(* IEC 61131-3 sources: station-control-three-platforms/codesys/src, 8 files *)

(* ---- ST_EvalRecipe.st ---- *)
// Evaluation recipe of FB_CurveEval as one structure. Not in the Siemens original: there the bench
// writes the recipe straight into the multi-instance Station.Eval. CODESYS refuses that
// (C0037 "'Eval' is no input of 'FB_HandleStation'"), so the station takes the recipe by reference
// and copies it into its own evaluation instance when it tares, once per part.
TYPE ST_EvalRecipe :
STRUCT
    Mode : INT := 3;
    GateX : REAL := 3.0;   // mm
    Gate2X : REAL := 10.0;   // mm
    PeakXLo : REAL := 13.0;   // mm
    PeakXHi : REAL := 26.0;   // mm
    StepSpan : REAL := 2.0;   // mm
    StopF : REAL := 30.0;   // N
    G1Lo : REAL;
    G1Hi : REAL;
    MeanLo : REAL;
    MeanHi : REAL;
    HystLo : REAL;
    HystHi : REAL;
    RetFMin : REAL;
    G2Lo : REAL;
    G2Hi : REAL;
    PeakFLo : REAL;
    PeakFHi : REAL;
    PeakXMin : REAL;
    PeakXMax : REAL;
    StepLo : REAL;
    StopXLo : REAL;
    StopXHi : REAL;
    EnvX0 : REAL := 1.0;   // mm
    EnvDx : REAL := 0.5;   // mm
    EnvN : INT := 55;
    EnvLo : ARRAY[0..63] OF REAL;   // N
    EnvHi : ARRAY[0..63] OF REAL;   // N
END_STRUCT
END_TYPE

(* ---- GVL_TestData.st ---- *)
// Generated by tools/testdata.py from siemens/scl/test/DB_TestData.scl. Do not edit.
// Recorded force-travel curves, the evaluation recipe and the expected values of the 14 replay cases.
{attribute 'qualified_only'}
VAR_GLOBAL
    NCurves : INT := 10;
    NCases : INT := 14;
    NSamples : INT := 5932;
    Tol : REAL := 0.001;
    GoodCurve : INT := 0;
    BadCurve : INT := 6;
    GateX : REAL := 3.0;
    Gate2X : REAL := 10.0;
    PeakXLo : REAL := 13.0;
    PeakXHi : REAL := 26.0;
    StepSpan : REAL := 2.0;
    StopF : REAL := 30.0;
    EnvX0 : REAL := 1.0;
    EnvDx : REAL := 0.5;
    EnvN : INT := 55;
    CurveStart : ARRAY[0..15] OF INT := [0, 620, 1246, 1746, 2366, 2988, 3606, 4228, 4728, 5310, 0, 0, 0, 0, 0, 0];
    CurveNPull : ARRAY[0..15] OF INT := [310, 313, 250, 310, 311, 309, 311, 250, 291, 311, 0, 0, 0, 0, 0, 0];
    CaseCurve : ARRAY[1..32] OF INT := [0, 1, 2, 3, 4, 5, 6, 7, 8, 9, 9, 8, 0, 3, 0, 0, 0, 0, 0, 0, 0, 0, 0, 0, 0, 0, 0, 0, 0, 0, 0, 0];
    CaseMode : ARRAY[1..32] OF INT := [3, 3, 3, 3, 3, 3, 3, 3, 3, 3, 2, 1, 4, 4, 0, 0, 0, 0, 0, 0, 0, 0, 0, 0, 0, 0, 0, 0, 0, 0, 0, 0];
    ExpOk : ARRAY[1..32] OF BOOL := [TRUE, TRUE, FALSE, FALSE, FALSE, FALSE, FALSE, FALSE, FALSE, FALSE, TRUE, TRUE, TRUE, TRUE, FALSE, FALSE, FALSE, FALSE, FALSE, FALSE, FALSE, FALSE, FALSE, FALSE, FALSE, FALSE, FALSE, FALSE, FALSE, FALSE, FALSE, FALSE];
    ExpNok : ARRAY[1..32] OF INT := [0, 0, 2, 2, 2, 3, 5, 2, 9, 2, 0, 0, 0, 0, 0, 0, 0, 0, 0, 0, 0, 0, 0, 0, 0, 0, 0, 0, 0, 0, 0, 0];
    ExpEnvViol : ARRAY[1..32] OF INT := [0, 0, 43, 0, 17, 41, 41, 43, 1, 0, 0, 1, 0, 0, 0, 0, 0, 0, 0, 0, 0, 0, 0, 0, 0, 0, 0, 0, 0, 0, 0, 0];
    ExpEnvNodes : ARRAY[1..32] OF INT := [55, 55, 46, 55, 55, 55, 55, 46, 55, 55, 55, 55, 55, 55, 0, 0, 0, 0, 0, 0, 0, 0, 0, 0, 0, 0, 0, 0, 0, 0, 0, 0];
    ExpFeat : ARRAY[0..287] OF REAL := [6.9821014, 5.37568, 6.1788907, 1.6064217, 10.845588, 16.818577, 19.848608, 3.9388027, 29.783041, 7.205183, 5.0210447, 6.113114, 2.1841383, 11.2528515, 17.15133, 18.303595, 4.152199, 30.096466, 4.183258, 2.565676, 3.374467, 1.6175817, 6.124597, 40.227142, 23.940363, 0.0, 23.785864, 5.1918726, 3.556863, 4.3743677, 1.6350094, 9.031395, 14.923322, 19.814, 3.9026327, 29.81065, 4.6947575, 3.0623243, 3.8785408, 1.632433, 8.425375, 14.073351, 19.786457, 3.8736982, 29.815647, 10.499536, 1.8700012, 6.184768, 8.629534, 14.390507, 20.330584, 19.78603, 3.8881645, 29.722036, 7.0127378, 5.3387175, 6.175728, 1.67402, 7.371472, 8.326099, 25.861488, 0.032551765, 29.877676, 4.238579, 2.6031868, 3.420883, 1.6353921, 6.187137, 41.858364, 23.904263, 0.0, 23.727392, 7.0128746, 5.3684235, 6.190649, 1.6444514, 10.856109, 16.749855, 19.791138, 3.8845482, 27.874788, 6.2380857, 2.573432, 4.405759, 3.6646535, 10.107543, 15.954138, 19.8363, 3.8773146, 29.792097, 6.2380857, 2.573432, 4.405759, 3.6646535, 10.107543, 15.954138, 19.8363, 3.8773146, 29.792097, 7.0128746, 5.3684235, 6.190649, 1.6444514, 10.856109, 16.749855, 19.791138, 3.8845482, 27.874788, 6.9821014, 5.37568, 6.1788907, 1.6064217, 10.845588, 16.818577, 19.848608, 3.9388027, 29.783041, 5.1918726, 3.556863, 4.3743677, 1.6350094, 9.031395, 14.923322, 19.814, 3.9026327, 29.81065, 0.0, 0.0, 0.0, 0.0, 0.0, 0.0, 0.0, 0.0, 0.0, 0.0, 0.0, 0.0, 0.0, 0.0, 0.0, 0.0, 0.0, 0.0, 0.0, 0.0, 0.0, 0.0, 0.0, 0.0, 0.0, 0.0, 0.0, 0.0, 0.0, 0.0, 0.0, 0.0, 0.0, 0.0, 0.0, 0.0, 0.0, 0.0, 0.0, 0.0, 0.0, 0.0, 0.0, 0.0, 0.0, 0.0, 0.0, 0.0, 0.0, 0.0, 0.0, 0.0, 0.0, 0.0, 0.0, 0.0, 0.0, 0.0, 0.0, 0.0, 0.0, 0.0, 0.0, 0.0, 0.0, 0.0, 0.0, 0.0, 0.0, 0.0, 0.0, 0.0, 0.0, 0.0, 0.0, 0.0, 0.0, 0.0, 0.0, 0.0, 0.0, 0.0, 0.0, 0.0, 0.0, 0.0, 0.0, 0.0, 0.0, 0.0, 0.0, 0.0, 0.0, 0.0, 0.0, 0.0, 0.0, 0.0, 0.0, 0.0, 0.0, 0.0, 0.0, 0.0, 0.0, 0.0, 0.0, 0.0, 0.0, 0.0, 0.0, 0.0, 0.0, 0.0, 0.0, 0.0, 0.0, 0.0, 0.0, 0.0, 0.0, 0.0, 0.0, 0.0, 0.0, 0.0, 0.0, 0.0, 0.0, 0.0, 0.0, 0.0, 0.0, 0.0, 0.0, 0.0, 0.0, 0.0, 0.0, 0.0, 0.0, 0.0, 0.0, 0.0, 0.0, 0.0, 0.0, 0.0, 0.0, 0.0, 0.0, 0.0, 0.0, 0.0, 0.0, 0.0, 0.0, 0.0, 0.0, 0.0, 0.0, 0.0];
    ExpFeatValid : ARRAY[0..287] OF BOOL := [TRUE, TRUE, TRUE, TRUE, TRUE, TRUE, TRUE, TRUE, TRUE, TRUE, TRUE, TRUE, TRUE, TRUE, TRUE, TRUE, TRUE, TRUE, TRUE, TRUE, TRUE, TRUE, TRUE, TRUE, TRUE, TRUE, TRUE, TRUE, TRUE, TRUE, TRUE, TRUE, TRUE, TRUE, TRUE, TRUE, TRUE, TRUE, TRUE, TRUE, TRUE, TRUE, TRUE, TRUE, TRUE, TRUE, TRUE, TRUE, TRUE, TRUE, TRUE, TRUE, TRUE, TRUE, TRUE, TRUE, TRUE, TRUE, TRUE, TRUE, TRUE, TRUE, TRUE, TRUE, TRUE, TRUE, TRUE, TRUE, TRUE, TRUE, TRUE, TRUE, TRUE, TRUE, TRUE, TRUE, TRUE, TRUE, TRUE, TRUE, TRUE, TRUE, TRUE, TRUE, TRUE, TRUE, TRUE, TRUE, TRUE, TRUE, TRUE, TRUE, TRUE, TRUE, TRUE, TRUE, TRUE, TRUE, TRUE, TRUE, TRUE, TRUE, TRUE, TRUE, TRUE, TRUE, TRUE, TRUE, TRUE, TRUE, TRUE, TRUE, TRUE, TRUE, TRUE, TRUE, TRUE, TRUE, TRUE, TRUE, TRUE, TRUE, TRUE, TRUE, TRUE, TRUE, FALSE, FALSE, FALSE, FALSE, FALSE, FALSE, FALSE, FALSE, FALSE, FALSE, FALSE, FALSE, FALSE, FALSE, FALSE, FALSE, FALSE, FALSE, FALSE, FALSE, FALSE, FALSE, FALSE, FALSE, FALSE, FALSE, FALSE, FALSE, FALSE, FALSE, FALSE, FALSE, FALSE, FALSE, FALSE, FALSE, FALSE, FALSE, FALSE, FALSE, FALSE, FALSE, FALSE, FALSE, FALSE, FALSE, FALSE, FALSE, FALSE, FALSE, FALSE, FALSE, FALSE, FALSE, FALSE, FALSE, FALSE, FALSE, FALSE, FALSE, FALSE, FALSE, FALSE, FALSE, FALSE, FALSE, FALSE, FALSE, FALSE, FALSE, FALSE, FALSE, FALSE, FALSE, FALSE, FALSE, FALSE, FALSE, FALSE, FALSE, FALSE, FALSE, FALSE, FALSE, FALSE, FALSE, FALSE, FALSE, FALSE, FALSE, FALSE, FALSE, FALSE, FALSE, FALSE, FALSE, FALSE, FALSE, FALSE, FALSE, FALSE, FALSE, FALSE, FALSE, FALSE, FALSE, FALSE, FALSE, FALSE, FALSE, FALSE, FALSE, FALSE, FALSE, FALSE, FALSE, FALSE, FALSE, FALSE, FALSE, FALSE, FALSE, FALSE, FALSE, FALSE, FALSE, FALSE, FALSE, FALSE, FALSE, FALSE, FALSE, FALSE, FALSE, FALSE, FALSE, FALSE, FALSE, FALSE, FALSE, FALSE, FALSE, FALSE, FALSE, FALSE, FALSE, FALSE, FALSE, FALSE, FALSE, FALSE, FALSE, FALSE, FALSE, FALSE, FALSE, FALSE, FALSE, FALSE, FALSE, FALSE, FALSE];
    Lim : ARRAY[0..63] OF REAL := [0.0, 0.0, 0.0, 0.0, 0.0, 0.0, 0.0, 0.0, 0.0, 15.241609, 18.417305, 0.0, 0.0, 0.0, 0.0, 0.0, 5.896105, 8.38203, 0.0, 0.0, 0.0, 0.0, 0.0, 9.4181, 12.402887, 14.982571, 18.676344, 17.139359, 22.516165, 2.9451215, 28.690018, 30.871372, 0.0, 0.0, 5.186474, 7.2080727, -0.5455249, 3.975223, 1.0, 9.212741, 12.608247, 14.728432, 18.930483, 16.769424, 22.886099, 2.8110514, 28.539938, 31.021452, 0.0, 0.0, 0.0, 0.0, 0.0, 0.0, 0.0, 0.0, 0.0, 0.0, 0.0, 0.0, 0.0, 0.0, 0.0, 0.0];
    EnvLo : ARRAY[0..63] OF REAL := [4.5024867, 4.5624857, 4.530773, 4.5635424, 4.573186, 4.617667, 4.6239376, 4.670679, 4.725596, 4.700003, 4.8820324, 4.926072, 5.163019, 5.6595745, 7.878658, 8.020163, 8.08159, 8.207902, 8.30263, 8.350869, 8.425625, 8.550419, 8.607436, 8.764787, 8.845735, 8.9147835, 8.99205, 9.068602, 9.331687, 9.416069, 9.513143, 9.665618, 10.123489, 10.642103, 11.14989, 11.027167, 10.830289, 10.428676, 10.27112, 10.313659, 10.363278, 10.468162, 10.585302, 10.677869, 10.748317, 10.8695135, 10.998811, 11.099038, 11.214338, 11.278554, 11.41541, 11.506263, 11.623229, 11.713954, 11.844806, 0.0, 0.0, 0.0, 0.0, 0.0, 0.0, 0.0, 0.0, 0.0];
    EnvHi : ARRAY[0..63] OF REAL := [9.917023, 9.98225, 9.992803, 10.004515, 10.029344, 10.026862, 10.070514, 10.102605, 12.041139, 12.557893, 12.779339, 12.91771, 13.360822, 13.471234, 13.533369, 13.642666, 13.729599, 13.860825, 13.911284, 13.990431, 14.0966015, 14.182879, 14.296827, 14.390328, 14.4539795, 14.551714, 14.698472, 15.185006, 15.688478, 16.23098, 16.795422, 17.309069, 17.854668, 18.362646, 18.931261, 18.921373, 19.396362, 19.986576, 19.496552, 19.897247, 19.346785, 18.766773, 16.553541, 16.354622, 16.457827, 16.512941, 16.617954, 16.769545, 16.847044, 16.997396, 17.054838, 17.213253, 17.348417, 17.397055, 17.536877, 0.0, 0.0, 0.0, 0.0, 0.0, 0.0, 0.0, 0.0, 0.0];
    X : ARRAY[0..5931] OF REAL := [0.0, -0.0033742767, 0.10472685, 0.19745024, 0.29981726, 0.39700347, 0.49491304, 0.6008226, 0.6972801, 0.7991843, 0.90281725, 0.99573755, 1.0995567, 1.1978173, 1.2951844, 1.3980939, 1.4998226, 1.5985514, 1.7018226, 1.8003706, 1.8912854, 1.999562, 2.0993705, 2.1909237, 2.2984662, 2.3891046, 2.4932854, 2.601009, 2.6959238, 2.796014, 2.894743, 2.9955568, 3.092743, 3.1978333, 3.292743, 3.3987377, 3.4987428, 3.59511, 3.6955674, 3.7989292, 3.8956633, 3.9927535, 4.0977483, 4.197296, 4.292573, 4.399477, 4.4931207, 4.593658, 4.6908493, 4.7944875, 4.8961205, 4.9969397, 5.094764, 5.18994, 5.2910357, 5.394844, 5.489573, 5.5893974, 5.6894984, 5.7891207, 5.893126, 5.989312, 6.076935, 6.1627493, 6.2443776, 6.328378, 6.4094586, 6.5168147, 6.6171765, 6.718815, 6.8094583, 6.9220915, 7.0171022, 7.1126394, 7.213565, 7.3112035, 7.4117403, 7.511751, 7.606661, 7.708384, 7.81248, 7.9090276, 8.005486, 8.110033, 8.2134, 8.307496, 8.410586, 8.505591, 8.600773, 8.702959, 8.809416, 8.908698, 8.999699, 9.103602, 9.201704, 9.301433, 9.39789, 9.503613, 9.601155, 9.699528, 9.802805, 9.89989, 10.003895, 10.098449, 10.201262, 10.298172, 10.399454, 10.497454, 10.592826, 10.699917, 10.798554, 10.89847, 10.996193, 11.098837, 11.192114, 11.287757, 11.391119, 11.496119, 11.592933, 11.693028, 11.786496, 11.891943, 11.991592, 12.0868635, 12.186582, 12.291321, 12.380411, 12.48514, 12.584327, 12.683965, 12.787603, 12.888337, 12.989885, 13.08306, 13.187704, 13.284523, 13.3848, 13.487896, 13.587353, 13.678811, 13.784454, 13.882715, 13.981008, 14.078545, 14.183087, 14.28164, 14.38038, 14.475013, 14.574927, 14.682922, 14.780104, 14.878199, 14.975023, 15.076039, 15.17287, 15.271434, 15.363907, 15.460098, 15.557104, 15.660487, 15.751045, 15.851062, 15.951705, 16.053541, 16.149647, 16.244019, 16.34385, 16.440685, 16.537062, 16.62862, 16.734083, 16.83637, 16.92229, 17.019585, 17.119505, 17.217972, 17.316803, 17.418, 17.508282, 17.611292, 17.70858, 17.800692, 17.902872, 17.99408, 18.09909, 18.191565, 18.287483, 18.387772, 18.49033, 18.585798, 18.676447, 18.777182, 18.874111, 18.979118, 19.070032, 19.165964, 19.270985, 19.360996, 19.462011, 19.55457, 19.65848, 19.755777, 19.848608, 19.970793, 20.087416, 20.211292, 20.32783, 20.445093, 20.557806, 20.648077, 20.741636, 20.84809, 20.953089, 21.043913, 21.147093, 21.24119, 21.348913, 21.449648, 21.545195, 21.634748, 21.745749, 21.841301, 21.946121, 22.040205, 22.143402, 22.240217, 22.341042, 22.44068, 22.53859, 22.634499, 22.738136, 22.838509, 22.941322, 23.042967, 23.129976, 23.239418, 23.335434, 23.430067, 23.531801, 23.641802, 23.734535, 23.835356, 23.933903, 24.02927, 24.133179, 24.232546, 24.332918, 24.43128, 24.52801, 24.624918, 24.728653, 24.823557, 24.925116, 25.026297, 25.123116, 25.230398, 25.325674, 25.426765, 25.523584, 25.621408, 25.71895, 25.820227, 25.919882, 26.019594, 26.116701, 26.216702, 26.315063, 26.42161, 26.524881, 26.622345, 26.714718, 26.815802, 26.917803, 27.014627, 27.115812, 27.214813, 27.312366, 27.413908, 27.51119, 27.612286, 27.709558, 27.811739, 27.911112, 28.007027, 28.111387, 28.199669, 28.301207, 28.40676, 28.508398, 28.60403, 28.701595, 28.8095, 28.900776, 29.00051, 29.101877, 29.200064, 29.301426, 29.398798, 29.500973, 29.572319, 29.6092, 29.646812, 29.686869, 29.716297, 29.758177, 29.799242, 29.837845, 29.867996, 29.91243, 29.94758, 29.943314, 29.928886, 29.886644, 29.850302, 29.813248, 29.77291, 29.739481, 29.693878, 29.666807, 29.625662, 29.588596, 29.545658, 29.446291, 29.346828, 29.248291, 29.144827, 29.049004, 28.937727, 28.847637, 28.75453, 28.642721, 28.549807, 28.448168, 28.348167, 28.251705, 28.151072, 28.05543, 27.9487, 27.857418, 27.751062, 27.654417, 27.556412, 27.45969, 27.360954, 27.257498, 27.15513, 27.059216, 26.958311, 26.85785, 26.761482, 26.654758, 26.5573, 26.460743, 26.360561, 26.257103, 26.160013, 26.06664, 25.96328, 25.863731, 25.76454, 25.668083, 25.56563, 25.464897, 25.367987, 25.26344, 25.167982, 25.070257, 24.966524, 24.871796, 24.767876, 24.67279, 24.576056, 24.471146, 24.368502, 24.26669, 24.170046, 24.073677, 23.97786, 23.87113, 23.777668, 23.676853, 23.576395, 23.480204, 23.375023, 23.272934, 23.17702, 23.081102, 22.978556, 22.88028, 22.779646, 22.677635, 22.582449, 22.482183, 22.376087, 22.28681, 22.185173, 22.084444, 21.981167, 21.891161, 21.780619, 21.684343, 21.589523, 21.48388, 21.391508, 21.285975, 21.187326, 21.08787, 20.986044, 20.88931, 20.790411, 20.692492, 20.591034, 20.4904, 20.394842, 20.293018, 20.197294, 20.102022, 19.994108, 19.893831, 19.797018, 19.694916, 19.590475, 19.501102, 19.397188, 19.298725, 19.19691, 19.100178, 18.99881, 18.902714, 18.797997, 18.700708, 18.604261, 18.502884, 18.39889, 18.303162, 18.206156, 18.103241, 17.99897, 17.907688, 17.802235, 17.704773, 17.608416, 17.508411, 17.407219, 17.30849, 17.209394, 17.109943, 17.011847, 16.906948, 16.809395, 16.708118, 16.613565, 16.507107, 16.412107, 16.31701, 16.208832, 16.112278, 16.011374, 15.918001, 15.814639, 15.7179, 15.617182, 15.515448, 15.413996, 15.3189, 15.21989, 15.117075, 15.018708, 14.91516, 14.81798, 14.721788, 14.619889, 14.519878, 14.4160595, 14.324873, 14.220602, 14.128693, 14.019857, 13.914687, 13.827314, 13.7215, 13.626677, 13.521501, 13.424581, 13.327847, 13.228756, 13.133394, 13.029112, 12.930293, 12.828841, 12.727287, 12.62883, 12.531464, 12.429921, 12.327181, 12.229639, 12.131453, 12.032723, 11.925458, 11.833815, 11.732442, 11.633894, 11.536803, 11.433075, 11.328346, 11.23716, 11.135245, 11.032245, 10.939425, 10.837878, 10.737963, 10.632873, 10.537234, 10.437139, 10.339868, 10.24041, 10.143681, 10.045037, 9.939037, 9.833128, 9.744676, 9.642303, 9.540303, 9.441941, 9.343032, 9.2415695, 9.141931, 9.047192, 8.943649, 8.843558, 8.747462, 8.645282, 8.554914, 8.446638, 8.344186, 8.247452, 8.145633, 8.051356, 7.9505424, 7.854803, 7.749255, 7.6534357, 7.5542603, 7.453893, 7.3493347, 7.2504253, 7.1519732, 7.054606, 6.9581485, 6.8538775, 6.7531433, 6.657409, 6.5563293, 6.4607816, 6.3632812, 6.274286, 6.1935673, 6.108753, 6.03021, 5.9339066, 5.8310876, 5.731545, 5.6369066, 5.531364, 5.437353, 5.337811, 5.2275395, 5.126901, 5.03872, 4.9384384, 4.8375287, 4.739082, 4.634901, 4.5331616, 4.4404383, 4.329167, 4.233348, 4.1344438, 4.0365286, 3.9392576, 3.834167, 3.7369862, 3.633433, 3.5345287, 3.4394383, 3.3372576, 3.2332575, 3.140433, 3.043066, 2.9320712, 2.8413372, 2.7396085, 2.6366086, 2.5347893, 2.441518, 2.342518, 2.2378001, 2.1382415, 2.034066, 1.9376031, 1.8358798, 1.7395127, 1.6385127, 1.540151, 1.4401511, 1.3368851, 1.2400553, 1.133151, 1.0449648, 0.939784, 0.8416882, 0.7337893, 0.6410499, 0.5402415, 0.43896484, 0.34032118, 0.23696484, 0.14223076, 0.03723076, 0.07943374, 0.0, 0.058969617, 0.1601451, 0.25842172, 0.36087385, 0.45877805, 0.5548792, 0.6574271, 0.75815046, 0.85487384, 0.9517888, 1.053975, 1.1582409, 1.2541559, 1.3572463, 1.4556025, 1.5523367, 1.6556187, 1.7556983, 1.8526186, 1.9547037, 2.0571558, 2.1517036, 2.2567995, 2.3577092, 2.4552517, 2.5556185, 2.6554377, 2.7547994, 2.850161, 2.9497144, 3.0517995, 3.1496186, 3.257076, 3.3558953, 3.4521666, 3.5518048, 3.653624, 3.7534378, 3.852991, 3.9552622, 4.04972, 4.1526294, 4.255996, 4.3528047, 4.4510016, 4.5480866, 4.6492677, 4.7482677, 4.853805, 4.9477253, 5.051906, 5.151358, 5.2348957, 5.3198113, 5.4007053, 5.4895253, 5.573419, 5.673228, 5.771866, 5.871143, 5.969329, 6.072978, 6.165616, 6.2763395, 6.37834, 6.4693394, 6.5714407, 6.6652493, 6.770627, 6.8630843, 6.9633555, 7.0697227, 7.168909, 7.2685523, 7.3637385, 7.4669037, 7.563648, 7.6645527, 7.7610154, 7.8674674, 7.9631057, 8.063478, 8.159749, 8.254574, 8.355664, 8.462856, 8.553574, 8.662393, 8.762766, 8.8588505, 8.952951, 9.056047, 9.15259, 9.251148, 9.357691, 9.453968, 9.555329, 9.654702, 9.75134, 9.855978, 9.954888, 10.04817, 10.15099, 10.252255, 10.3547125, 10.451904, 10.551271, 10.646809, 10.748909, 10.853186, 10.952457, 11.050553, 11.14801, 11.246378, 11.350468, 11.444835, 11.546383, 11.644745, 11.748659, 11.844665, 11.942393, 12.038213, 12.13958, 12.245122, 12.339048, 12.439409, 12.540957, 12.639862, 12.740053, 12.837516, 12.932607, 13.040059, 13.139059, 13.238154, 13.338431, 13.4359, 13.5304575, 13.635559, 13.72675, 13.818857, 13.918681, 14.016246, 14.117352, 14.217459, 14.311023, 14.407762, 14.50431, 14.610332, 14.701975, 14.796544, 14.899007, 14.994475, 15.085858, 15.194316, 15.28988, 15.3827095, 15.478273, 15.579289, 15.676763, 15.776773, 15.875156, 15.973704, 16.068811, 16.163736, 16.2553, 16.359764, 16.457323, 16.552242, 16.653168, 16.743004, 16.841015, 16.939758, 17.037136, 17.140327, 17.235802, 17.331541, 17.428104, 17.52593, 17.631126, 17.718876, 17.81943, 17.915802, 18.00819, 18.111834, 18.202488, 18.303595, 18.407286, 18.52944, 18.65905, 18.7763, 18.901001, 19.0094, 19.106045, 19.20614, 19.303415, 19.40779, 19.507235, 19.609697, 19.70224, 19.802341, 19.900156, 20.002895, 20.102533, 20.202618, 20.304895, 20.402363, 20.497267, 20.599997, 20.69355, 20.796188, 20.893097, 20.992193, 21.097012, 21.191204, 21.29547, 21.400927, 21.492119, 21.598661, 21.689854, 21.794113, 21.885592, 21.988316, 22.08878, 22.190773, 22.293049, 22.38805, 22.484604, 22.585506, 22.687784, 22.784433, 22.885614, 22.98833, 23.082354, 23.185162, 23.283348, 23.381716, 23.482725, 23.583992, 23.68372, 23.78337, 23.879997, 23.972647, 24.07764, 24.179012, 24.279741, 24.376842, 24.48021, 24.577572, 24.6793, 24.773943, 24.874945, 24.974407, 25.07404, 25.175955, 25.274588, 25.366964, 25.468056, 25.566055, 25.66897, 25.770609, 25.869247, 25.965885, 26.0708, 26.170258, 26.2708, 26.36344, 26.460264, 26.56645, 26.666822, 26.763725, 26.867178, 26.958647, 27.05411, 27.163929, 27.263475, 27.364023, 27.460024, 27.559578, 27.659397, 27.761215, 27.85913, 27.956684, 28.054413, 28.157417, 28.249779, 28.357328, 28.453423, 28.551237, 28.653881, 28.746983, 28.850885, 28.955158, 29.047626, 29.149813, 29.249632, 29.350636, 29.44836, 29.546822, 29.64455, 29.74519, 29.845291, 29.898531, 29.932146, 29.975742, 30.014538, 30.052784, 30.09384, 30.124363, 30.161966, 30.199852, 30.23428, 30.276073, 30.279707, 30.259258, 30.220552, 30.182497, 30.147161, 30.109282, 30.07712, 30.027245, 29.995913, 29.958479, 29.921057, 29.88163, 29.803432, 29.702337, 29.604788, 29.508512, 29.404512, 29.309692, 29.208055, 29.105412, 29.010315, 28.907495, 28.810219, 28.708496, 28.606033, 28.511213, 28.409018, 28.308836, 28.206108, 28.11083, 28.009554, 27.920464, 27.817097, 27.714096, 27.614098, 27.519081, 27.421623, 27.311539, 27.215809, 27.113165, 27.011442, 26.923613, 26.819523, 26.72316, 26.624512, 26.518154, 26.424501, 26.324501, 26.223682, 26.12832, 26.023682, 25.925581, 25.826756, 25.725304, 25.633213, 25.526209, 25.431484, 25.327932, 25.231379, 25.124107, 25.027378, 24.92774, 24.827005, 24.72682, 24.634266, 24.533634, 24.435629, 24.333357, 24.235714, 24.134075, 24.037159, 23.934883, 23.83689, 23.733522, 23.644058, 23.538336, 23.439335, 23.337143, 23.241873, 23.141325, 23.039495, 22.943308, 22.836676, 22.740585, 22.643122, 22.548845, 22.443756, 22.34893, 22.245022, 22.14148, 22.045925, 21.948095, 21.845825, 21.747463, 21.648638, 21.544724, 21.452633, 21.34591, 21.252352, 21.149809, 21.053707, 20.957075, 20.850708, 20.75434, 20.64933, 20.556244, 20.450605, 20.35551, 20.255686, 20.158957, 20.061596, 19.960772, 19.857952, 19.762127, 19.659489, 19.561398, 19.463669, 19.359297, 19.259573, 19.161749, 19.060844, 18.962467, 18.862371, 18.765282, 18.660913, 18.566366, 18.460653, 18.360914, 18.270807, 18.172451, 18.065079, 17.969627, 17.871622, 17.768164, 17.67243, 17.567436, 17.47643, 17.368792, 17.271786, 17.17751, 17.071148, 16.969872, 16.872866, 16.770239, 16.681765, 16.574047, 16.477217, 16.370668, 16.275764, 16.177212, 16.073658, 15.979759, 15.87902, 15.777563, 15.671382, 15.586376, 15.481924, 15.379919, 15.276377, 15.181281, 15.08636, 14.982185, 14.887541, 14.778909, 14.685083, 14.590627, 14.482345, 14.385892, 14.288073, 14.186977, 14.087796, 13.983977, 13.882429, 13.788419, 13.691237, 13.585786, 13.489599, 13.390775, 13.289956, 13.196493, 13.09286, 12.993312, 12.887945, 12.791126, 12.695663, 12.598573, 12.4952965, 12.398929, 12.295924, 12.19511, 12.095748, 11.997562, 11.899285, 11.795099, 11.700924, 11.59928, 11.501275, 11.400998, 11.296269, 11.20136, 11.098631, 10.997439, 10.901258, 10.802343, 10.704705, 10.604073, 10.503344, 10.405062, 10.304508, 10.20687, 10.110237, 10.015503, 9.908232, 9.80387, 9.70986, 9.613317, 9.510488, 9.412759, 9.315125, 9.2118435, 9.115025, 9.007386, 8.917743, 8.812657, 8.711567, 8.614014, 8.5132, 8.413094, 8.316461, 8.2181835, 8.115466, 8.0167265, 7.91754, 7.821811, 7.720806, 7.614529, 7.5185294, 7.415439, 7.320343, 7.2262526, 7.1214337, 7.015976, 6.92479, 6.824875, 6.7247844, 6.624508, 6.5194283, 6.4205985, 6.325327, 6.2258644, 6.1244917, 6.02304, 5.9274974, 5.825758, 5.7219496, 5.6314015, 5.536194, 5.44547, 5.3669214, 5.285751, 5.202383, 5.105436, 5.006702, 4.9036064, 4.806521, 4.706877, 4.6049786, 4.5074253, 4.4004254, 4.30834, 4.207973, 4.1086006, 4.004883, 3.9012392, 3.8079624, 3.7125103, 3.6096008, 3.5041487, 3.413053, 3.30342, 3.21142, 3.1053243, 3.0126913, 2.9129572, 2.8093243, 2.699053, 2.6135051, 2.506138, 2.4069571, 2.3082337, 2.2100475, 2.1109626, 2.00642, 1.910505, 1.8110476, 1.7060529, 1.6115955, 1.5136752, 1.4113135, 1.3050423, 1.2158561, 1.1087602, 1.0117602, 0.9073135, 0.8141273, 0.7076752, 0.6063986, 0.50649434, 0.40968055, 0.31476563, 0.20966984, 0.11121774, 0.008217737, 0.0, 0.08626114, 0.16408622, 0.25262398, 0.34693274, 0.44683695, 0.5450178, 0.64548063, 0.7489327, 0.841486, 0.944571, 1.047401, 1.1493956, 1.2461296, 1.3409435, 1.4471296, 1.5429435, 1.6451297, 1.7413158, 1.8395978, 1.9470446, 2.046316, 2.141688, 2.2395074, 2.3439596, 2.440784, 2.540598, 2.6418743, 2.7417786, 2.8391511, 2.9425128, 3.0404222, 3.1325235, 3.2412467, 3.3387947, 3.4342575, 3.5342574, 3.6396246, 3.7380767, 3.8398108, 3.9381723, 4.034534, 4.13063, 4.2379065, 4.332268, 4.4399066, 4.5368214, 4.628816, 4.735364, 4.836087, 4.928742, 5.0387416, 5.130109, 5.239098, 5.3370132, 5.43438, 5.5339227, 5.6311035, 5.731024, 5.8305664, 5.924747, 6.027933, 6.1294813, 6.2354865, 6.3234863, 6.43004, 6.530306, 6.6274014, 6.7249546, 6.8309493, 6.9234123, 7.0274973, 7.1264067, 7.2263165, 7.329322, 7.422141, 7.5283217, 7.6280613, 7.7241464, 7.820609, 7.923875, 8.022885, 8.123976, 8.231061, 8.323157, 8.426066, 8.522167, 8.62453, 8.719806, 8.822077, 8.918812, 9.018099, 9.116663, 9.21195, 9.308865, 9.403785, 9.504344, 9.603817, 9.694104, 9.796387, 9.90503, 9.994046, 10.088147, 10.185254, 10.283903, 10.380095, 10.480473, 10.572754, 10.679222, 10.772696, 10.870611, 10.970898, 11.067276, 11.16219, 11.261116, 11.365132, 11.458878, 11.550426, 11.658532, 11.751276, 11.844559, 11.944931, 12.048128, 12.144404, 12.240521, 12.341804, 12.436001, 12.537735, 12.632028, 12.722315, 12.822873, 12.918155, 13.020804, 13.11182, 13.215831, 13.312203, 13.411315, 13.506406, 13.602703, 13.704895, 13.813751, 13.936825, 14.052898, 14.177792, 14.293041, 14.399817, 14.500093, 14.601089, 14.699647, 14.798828, 14.900009, 14.99928, 15.095919, 15.194653, 15.2962055, 15.402014, 15.493297, 15.597206, 15.696291, 15.793211, 15.894573, 15.994216, 16.094482, 16.197584, 16.296854, 16.395493, 16.494854, 16.593866, 16.69186, 16.793776, 16.89269, 16.994047, 17.094774, 17.193243, 17.292328, 17.389967, 17.489605, 17.591696, 17.690153, 17.79379, 17.88644, 17.984615, 18.091429, 18.188078, 18.289797, 18.389711, 18.487074, 18.585089, 18.683716, 18.787716, 18.88736, 18.982813, 19.084908, 19.180637, 19.287733, 19.378914, 19.481653, 19.58519, 19.688015, 19.784105, 19.885105, 19.981941, 20.080477, 20.177025, 20.277748, 20.381495, 20.474669, 20.585121, 20.684946, 20.782211, 20.869228, 20.983856, 21.075409, 21.175041, 21.27759, 21.37559, 21.48168, 21.57587, 21.669786, 21.769611, 21.87778, 21.970972, 22.07425, 22.1737, 22.27034, 22.372978, 22.464525, 22.568436, 22.673801, 22.76935, 22.873451, 22.968447, 23.068174, 23.167181, 23.262638, 23.363457, 23.448547, 23.490519, 23.525759, 23.558645, 23.595072, 23.638952, 23.6792, 23.715626, 23.748682, 23.789104, 23.828627, 23.864237, 23.902477, 23.940363, 23.9459, 23.91903, 23.88006, 23.848814, 23.799929, 23.76615, 23.732264, 23.693836, 23.654856, 23.61289, 23.575373, 23.54095, 23.499975, 23.465818, 23.40177, 23.306679, 23.211945, 23.113216, 23.009312, 22.915482, 22.810843, 22.714844, 22.607939, 22.5082, 22.41111, 22.315023, 22.216562, 22.114561, 22.017641, 21.91356, 21.818556, 21.71846, 21.61546, 21.519827, 21.423178, 21.322727, 21.2219, 21.118635, 21.017353, 20.921162, 20.821173, 20.717806, 20.617353, 20.519167, 20.423529, 20.323885, 20.222248, 20.122982, 20.017609, 19.922152, 19.82279, 19.728874, 19.628683, 19.527231, 19.420507, 19.328598, 19.226055, 19.12614, 19.027859, 18.92413, 18.830034, 18.725492, 18.621853, 18.528305, 18.429848, 18.329391, 18.231758, 18.133385, 18.02812, 17.93539, 17.828562, 17.731556, 17.632019, 17.53247, 17.435652, 17.331741, 17.23164, 17.13119, 17.039188, 16.934822, 16.834013, 16.72946, 16.632635, 16.541449, 16.433624, 16.337263, 16.238619, 16.140078, 16.041264, 15.936167, 15.837439, 15.731354, 15.643433, 15.542253, 15.437524, 15.340157, 15.234438, 15.1426935, 15.038332, 14.945151, 14.839055, 14.736237, 14.64305, 14.54605, 14.445321, 14.343502, 14.241587, 14.14296, 14.043225, 13.940954, 13.848028, 13.748943, 13.649853, 13.5404005, 13.445395, 13.346565, 13.251119, 13.149114, 13.047938, 12.949023, 12.845475, 12.744108, 12.648922, 12.546831, 12.443922, 12.351374, 12.2532835, 12.144917, 12.04564, 11.948273, 11.850539, 11.755182, 11.652087, 11.552539, 11.4536295, 11.353901, 11.25381, 11.150906, 11.051443, 10.959076, 10.856342, 10.759076, 10.655523, 10.555251, 10.460879, 10.356331, 10.25497, 10.159789, 10.060602, 9.955512, 9.858231, 9.758411, 9.658512, 9.55823, 9.461773, 9.35714, 9.258135, 9.159677, 9.060767, 8.962858, 8.86222, 8.762124, 8.663587, 8.565485, 8.465938, 8.362666, 8.270204, 8.161209, 8.063927, 7.969384, 7.865379, 7.757927, 7.661746, 7.571554, 7.4681025, 7.373012, 7.262645, 7.166826, 7.067826, 6.965905, 6.872453, 6.765549, 6.6689053, 6.567815, 6.467815, 6.374448, 6.27481, 6.170256, 6.0742564, 5.970443, 5.867533, 5.775799, 5.669251, 5.576607, 5.4744263, 5.37507, 5.274251, 5.173602, 5.0736976, 4.973969, 4.87824, 4.7821445, 4.680597, 4.5706925, 4.4696817, 4.3800435, 4.268049, 4.172134, 4.080586, 3.9725008, 3.8796763, 3.7860382, 3.6812189, 3.5841231, 3.479304, 3.376038, 3.285123, 3.1766655, 3.0816603, 2.9889317, 2.8742027, 2.7805698, 2.6814742, 2.58474, 2.4808357, 2.3843784, 2.2894688, 2.1821017, 2.0858252, 1.9848198, 1.8824581, 1.7823783, 1.689091, 1.5809155, 1.4890857, 1.3824581, 1.2849952, 1.1856335, 1.0859048, 0.9898941, 0.8930803, 0.7830696, 0.6876282, 0.5891654, 0.48952705, 0.39324507, 0.29234084, 0.20517014, 0.11862703, 0.044536024, 0.0, 0.059942853, 0.15758651, 0.25440568, 0.3589482, 0.46004933, 0.5611344, 0.6548631, 0.75676733, 0.86150146, 0.95358115, 1.0613099, 1.1569589, 1.2548631, 1.3582249, 1.4564961, 1.5571398, 1.6575068, 1.7561344, 1.8561398, 1.9555973, 2.055959, 2.15731, 2.2549536, 2.355693, 2.4565973, 2.5547833, 2.653778, 2.7529643, 2.8573205, 2.9499643, 3.0485973, 3.154326, 3.258145, 3.3519697, 3.4530602, 3.5616877, 3.6537888, 3.7530653, 3.8539696, 3.9496984, 4.048975, 4.15506, 4.2600656, 4.3559694, 4.450241, 4.553613, 4.6583314, 4.7553368, 4.8541613, 4.952624, 5.0506186, 5.1556134, 5.2568846, 5.3572516, 5.4571557, 5.5487146, 5.6542516, 5.7500815, 5.848257, 5.946342, 6.0442944, 6.131662, 6.2118382, 6.2960143, 6.375015, 6.475398, 6.5699406, 6.673946, 6.7746744, 6.876488, 6.9773183, 7.0665946, 7.1729617, 7.27168, 7.3722386, 7.4740577, 7.5736055, 7.6791425, 7.767797, 7.8653398, 7.969797, 8.065621, 8.167153, 8.269989, 8.361536, 8.461175, 8.568446, 8.663994, 8.763, 8.869728, 8.967185, 9.065, 9.166371, 9.254648, 9.360101, 9.46093, 9.563106, 9.661111, 9.7617445, 9.856659, 9.962297, 10.057298, 10.164111, 10.258941, 10.361484, 10.453223, 10.551409, 10.659042, 10.756239, 10.855047, 10.954414, 11.057234, 11.149872, 11.254872, 11.352612, 11.447612, 11.55634, 11.652515, 11.749978, 11.846899, 11.953888, 12.050718, 12.148436, 12.250532, 12.347176, 12.448813, 12.549452, 12.646452, 12.7430105, 12.8481865, 12.946457, 13.047372, 13.147378, 13.250473, 13.3443775, 13.441564, 13.545021, 13.642846, 13.746388, 13.845665, 13.943575, 14.038495, 14.137947, 14.241128, 14.341495, 14.437409, 14.545048, 14.636771, 14.736697, 14.835883, 14.933149, 15.03534, 15.131453, 15.23091, 15.330197, 15.4204, 15.52323, 15.6187935, 15.709166, 15.815352, 15.914922, 16.00639, 16.110039, 16.208954, 16.302608, 16.396261, 16.497183, 16.591007, 16.693203, 16.793215, 16.88896, 16.986065, 17.089806, 17.184998, 17.2752, 17.376476, 17.468401, 17.57196, 17.669874, 17.769077, 17.861189, 17.959019, 18.059114, 18.161945, 18.251875, 18.350977, 18.449902, 18.548456, 18.64293, 18.740578, 18.837872, 18.937328, 19.02971, 19.129723, 19.232094, 19.325014, 19.422764, 19.525595, 19.613792, 19.719078, 19.814, 19.919504, 20.04212, 20.15819, 20.281082, 20.401524, 20.511564, 20.60375, 20.707033, 20.808395, 20.91049, 21.010033, 21.10931, 21.2064, 21.304592, 21.406315, 21.508495, 21.6065, 21.704512, 21.798693, 21.906687, 21.997974, 22.100151, 22.204704, 22.302252, 22.39762, 22.504076, 22.600353, 22.696167, 22.79672, 22.903719, 22.993368, 23.094183, 23.198092, 23.299007, 23.396645, 23.495646, 23.593475, 23.692747, 23.791107, 23.893204, 23.99648, 24.092756, 24.191118, 24.289673, 24.395853, 24.491858, 24.584322, 24.686327, 24.790226, 24.88778, 24.98996, 25.084875, 25.183603, 25.28597, 25.391157, 25.48106, 25.583986, 25.681438, 25.78654, 25.882534, 25.976997, 26.084625, 26.178997, 26.279093, 26.380821, 26.480001, 26.584827, 26.674923, 26.775928, 26.882019, 26.97811, 27.076385, 27.172386, 27.27448, 27.374933, 27.473944, 27.57186, 27.674858, 27.774858, 27.871407, 27.970226, 28.07169, 28.170599, 28.272417, 28.366512, 28.4667, 28.564981, 28.665806, 28.770975, 28.865072, 28.963987, 29.059992, 29.169172, 29.265812, 29.362364, 29.462551, 29.55378, 29.593468, 29.635618, 29.666414, 29.698565, 29.740263, 29.778048, 29.8223, 29.86127, 29.90024, 29.936306, 29.971361, 29.971085, 29.944763, 29.909967, 29.872366, 29.835667, 29.80542, 29.759996, 29.717112, 29.685328, 29.645077, 29.608839, 29.573593, 29.501139, 29.405039, 29.305681, 29.206215, 29.103575, 29.009033, 28.904667, 28.804937, 28.710293, 28.605474, 28.508661, 28.417282, 28.311565, 28.214464, 28.114277, 28.012548, 27.913092, 27.820448, 27.71899, 27.618353, 27.514618, 27.415438, 27.320534, 27.218431, 27.11598, 27.018234, 26.922245, 26.822065, 26.722776, 26.62123, 26.523596, 26.426495, 26.323044, 26.222862, 26.12549, 26.024942, 25.92758, 25.820772, 25.725574, 25.629202, 25.528017, 25.425926, 25.324293, 25.22792, 25.126825, 25.029005, 24.933367, 24.829548, 24.730543, 24.63091, 24.531271, 24.427984, 24.337261, 24.231985, 24.136707, 24.031889, 23.931883, 23.831882, 23.73997, 23.641516, 23.532425, 23.435963, 23.343596, 23.237778, 23.142862, 23.039133, 22.941957, 22.839037, 22.74458, 22.63958, 22.542213, 22.444937, 22.347937, 22.243298, 22.14175, 22.049746, 21.94365, 21.849377, 21.7401, 21.650915, 21.54883, 21.443733, 21.34736, 21.248903, 21.14999, 21.053713, 20.948261, 20.850527, 20.752527, 20.654068, 20.551973, 20.450611, 20.353426, 20.247616, 20.158962, 20.056686, 19.95451, 19.848787, 19.76441, 19.6565, 19.555319, 19.45823, 19.358404, 19.264393, 19.158207, 19.05784, 18.959488, 18.859291, 18.76084, 18.65584, 18.561293, 18.458387, 18.365738, 18.261276, 18.16474, 18.065456, 17.959185, 17.868, 17.770355, 17.661999, 17.565441, 17.466255, 17.363897, 17.270435, 17.170887, 17.071249, 16.968435, 16.872057, 16.771149, 16.675966, 16.571058, 16.47269, 16.371775, 16.271776, 16.172047, 16.071234, 15.967866, 15.878132, 15.776042, 15.676312, 15.57985, 15.473297, 15.378382, 15.279025, 15.177201, 15.079201, 14.981653, 14.875744, 14.789733, 14.678914, 14.583095, 14.475462, 14.384275, 14.279727, 14.186456, 14.079722, 13.987535, 13.88844, 13.783078, 13.69144, 13.58844, 13.489435, 13.387791, 13.282164, 13.192785, 13.088605, 12.986334, 12.884238, 12.789509, 12.687323, 12.587961, 12.48569, 12.391137, 12.28995, 12.1933975, 12.090126, 11.99194, 11.893216, 11.788483, 11.695754, 11.591849, 11.499387, 11.3926525, 11.294375, 11.194839, 11.092557, 10.997738, 10.890556, 10.798822, 10.69428, 10.595455, 10.501907, 10.401269, 10.301546, 10.204168, 10.10453, 9.9986315, 9.900072, 9.803525, 9.699344, 9.605338, 9.499519, 9.406876, 9.300428, 9.201333, 9.105418, 9.001323, 8.907136, 8.802052, 8.707588, 8.607865, 8.513311, 8.412035, 8.308216, 8.204583, 8.110939, 8.007684, 7.9073915, 7.813301, 7.709386, 7.6157475, 7.509753, 7.409833, 7.307189, 7.2156467, 7.115641, 7.0119123, 6.9109178, 6.8138165, 6.7170825, 6.618269, 6.5197263, 6.416269, 6.3316565, 6.241204, 6.1591926, 6.0856547, 5.9944844, 5.894399, 5.7966704, 5.6911173, 5.593761, 5.493942, 5.3995748, 5.2914844, 5.1911173, 5.095665, 4.987128, 4.8909416, 4.793027, 4.6963882, 4.5995693, 4.4999366, 4.4001174, 4.2952023, 4.1964736, 4.096298, 4.002112, 3.892383, 3.7965639, 3.6973832, 3.596197, 3.495383, 3.3942926, 3.2942874, 3.1958299, 3.094931, 2.997197, 2.8948298, 2.7965586, 2.6989202, 2.597463, 2.494101, 2.3953724, 2.299649, 2.196016, 2.1035533, 2.0005586, 1.9009149, 1.7969257, 1.702282, 1.5964628, 1.5001011, 1.3938245, 1.3030107, 1.1989149, 1.0978192, 0.99527663, 0.89845747, 0.8009096, 0.6996383, 0.60026056, 0.50273407, 0.39791492, 0.29663295, 0.20254253, 0.10845211, -0.0033723959, 0.0, 0.025911892, 0.12764062, 0.2301778, 0.32582146, 0.42782146, 0.5292682, 0.6247364, 0.7245502, 0.82582146, 0.9259119, 1.0321778, 1.1327311, 1.2300928, 1.3288268, 1.4261938, 1.524731, 1.6241832, 1.7260131, 1.8231034, 1.9323747, 2.026098, 2.1261885, 2.2300076, 2.326013, 2.429545, 2.5251832, 2.626465, 2.7291992, 2.82646, 2.9284651, 3.0237417, 3.1271088, 3.2188323, 3.3277419, 3.4281034, 3.5262842, 3.6254652, 3.7312844, 3.8243802, 3.9309225, 4.0269175, 4.123109, 4.223928, 4.3228374, 4.425109, 4.525572, 4.6247525, 4.7195716, 4.822114, 4.9290237, 5.0293, 5.1238375, 5.2208376, 5.3288484, 5.4212046, 5.5208535, 5.6197524, 5.7191143, 5.8213906, 5.91721, 6.024593, 6.099498, 6.184956, 6.2723126, 6.350122, 6.4428988, 6.5479894, 6.6529894, 6.745814, 6.8487177, 6.9472713, 7.035271, 7.144271, 7.238819, 7.341181, 7.4426327, 7.544372, 7.642824, 7.739106, 7.842649, 7.943654, 8.03675, 8.132574, 8.232659, 8.330755, 8.439484, 8.538937, 8.632404, 8.740123, 8.838304, 8.93659, 9.036857, 9.1335, 9.236138, 9.329867, 9.441229, 9.532867, 9.63041, 9.731968, 9.836782, 9.934687, 10.030703, 10.1319685, 10.225612, 10.330792, 10.433166, 10.529888, 10.630798, 10.730081, 10.825798, 10.926899, 11.02517, 11.123815, 11.225634, 11.326186, 11.426543, 11.529186, 11.621825, 11.720729, 11.820463, 11.919373, 12.023655, 12.127926, 12.2206545, 12.318564, 12.427474, 12.514117, 12.62366, 12.719671, 12.820032, 12.917038, 13.015592, 13.123953, 13.222676, 13.317947, 13.420511, 13.5199585, 13.618325, 13.716778, 13.815873, 13.913511, 14.017325, 14.120155, 14.219336, 14.318698, 14.4135275, 14.515794, 14.611895, 14.711171, 14.814623, 14.910176, 15.008724, 15.108283, 15.208299, 15.299219, 15.397868, 15.499246, 15.597528, 15.69463, 15.784826, 15.888932, 15.987401, 16.084778, 16.17688, 16.277077, 16.375822, 16.474646, 16.573385, 16.667673, 16.769327, 16.866146, 16.960077, 17.057093, 17.158833, 17.259024, 17.352764, 17.458775, 17.544249, 17.644077, 17.743546, 17.84147, 17.936115, 18.032679, 18.130865, 18.22634, 18.327354, 18.425455, 18.527014, 18.623207, 18.719685, 18.813051, 18.916706, 19.010988, 19.104372, 19.19511, 19.297031, 19.396318, 19.499786, 19.601984, 19.691265, 19.786457, 19.895712, 20.013876, 20.135775, 20.25421, 20.382725, 20.4863, 20.591118, 20.683401, 20.788671, 20.885853, 20.984491, 21.08622, 21.181225, 21.282236, 21.384502, 21.48114, 21.588694, 21.678518, 21.781065, 21.880337, 21.975891, 22.07916, 22.182253, 22.2738, 22.384077, 22.48172, 22.582172, 22.679268, 22.774448, 22.880901, 22.972816, 23.07282, 23.175104, 23.271093, 23.370188, 23.478651, 23.57511, 23.670933, 23.773375, 23.874746, 23.974922, 24.07039, 24.167843, 24.270939, 24.375843, 24.473125, 24.571033, 24.666588, 24.763412, 24.86614, 24.969322, 25.059864, 25.162874, 25.268332, 25.369146, 25.4637, 25.556253, 25.663433, 25.759253, 25.857885, 25.96253, 26.060162, 26.153727, 26.260992, 26.36054, 26.461449, 26.56745, 26.662998, 26.755919, 26.854195, 26.961098, 27.058743, 27.158104, 27.25302, 27.356295, 27.460752, 27.554663, 27.651747, 27.752583, 27.850763, 27.956583, 28.05231, 28.153673, 28.251131, 28.347227, 28.45305, 28.550322, 28.644514, 28.746424, 28.850885, 28.945429, 29.045786, 29.144157, 29.248976, 29.344795, 29.447987, 29.54119, 29.580042, 29.62329, 29.656717, 29.69505, 29.733934, 29.772356, 29.803427, 29.852116, 29.881182, 29.923882, 29.96567, 29.996645, 29.996737, 29.976862, 29.937529, 29.899372, 29.862036, 29.82715, 29.790722, 29.751476, 29.716873, 29.671541, 29.637661, 29.600325, 29.562891, 29.493938, 29.387024, 29.2883, 29.18838, 29.090826, 28.990469, 28.890465, 28.78956, 28.687284, 28.590454, 28.49291, 28.390278, 28.291086, 28.196081, 28.096172, 27.991726, 27.88872, 27.7918, 27.692528, 27.598162, 27.50016, 27.389433, 27.29598, 27.19614, 27.10115, 26.999146, 26.898874, 26.802326, 26.699778, 26.604502, 26.505587, 26.398949, 26.30531, 26.21257, 26.1043, 26.00357, 25.900293, 25.804028, 25.70066, 25.603289, 25.501745, 25.402836, 25.309374, 25.207277, 25.106554, 25.017906, 24.908, 24.813635, 24.711176, 24.607452, 24.511442, 24.411905, 24.309532, 24.210623, 24.106895, 24.011885, 23.915064, 23.817879, 23.718336, 23.612879, 23.512873, 23.41915, 23.316235, 23.218868, 23.11732, 23.018139, 22.920315, 22.81941, 22.722948, 22.620123, 22.517574, 22.420574, 22.315123, 22.222755, 22.12566, 22.023117, 21.925192, 21.825563, 21.73065, 21.628372, 21.526367, 21.430271, 21.318914, 21.221, 21.128363, 21.02709, 20.929272, 20.824905, 20.726627, 20.62608, 20.528803, 20.428804, 20.329521, 20.232985, 20.126698, 20.030516, 19.936245, 19.833143, 19.73016, 19.634686, 19.531963, 19.437681, 19.332415, 19.23041, 19.130772, 19.034128, 18.935862, 18.835857, 18.7344, 18.637123, 18.539303, 18.435846, 18.342299, 18.23548, 18.132648, 18.038568, 17.937197, 17.84265, 17.740011, 17.6401, 17.539553, 17.443005, 17.345728, 17.248362, 17.139723, 17.042265, 16.949175, 16.84508, 16.7459, 16.651165, 16.548887, 16.443527, 16.346441, 16.250431, 16.14734, 16.052414, 15.950516, 15.8478775, 15.748414, 15.6508665, 15.549968, 15.453686, 15.353233, 15.2566805, 15.15468, 15.050313, 14.949765, 14.850856, 14.756941, 14.651936, 14.55458, 14.456659, 14.354032, 14.254026, 14.164557, 14.057015, 13.9621, 13.859839, 13.757015, 13.659914, 13.562005, 13.460457, 13.358547, 13.261728, 13.160632, 13.05718, 12.960356, 12.859446, 12.753175, 12.659808, 12.562978, 12.462707, 12.362706, 12.260882, 12.162425, 12.066069, 11.965696, 11.861158, 11.766967, 11.663696, 11.5686, 11.47168, 11.362696, 11.268866, 11.17177, 11.066137, 10.965228, 10.866946, 10.769228, 10.670036, 10.572036, 10.473488, 10.372393, 10.273207, 10.173297, 10.077653, 9.974563, 9.869749, 9.773738, 9.665658, 9.570834, 9.477557, 9.377461, 9.272547, 9.181094, 9.080542, 8.974089, 8.876733, 8.78218, 8.680536, 8.580536, 8.477078, 8.378435, 8.278711, 8.181706, 8.077887, 7.98052, 7.883791, 7.7804294, 7.676073, 7.583424, 7.4855146, 7.3815036, 7.286509, 7.1853228, 7.087509, 6.980594, 6.885408, 6.786227, 6.686775, 6.5914025, 6.4840407, 6.388397, 6.300397, 6.2213163, 6.139406, 6.047693, 5.965804, 5.8651657, 5.7661657, 5.66598, 5.567799, 5.463437, 5.359437, 5.2632565, 5.167432, 5.0657086, 4.9659796, 4.869437, 4.767799, 4.6630754, 4.566336, 4.463347, 4.3684425, 4.268799, 4.167703, 4.0643415, 3.9627085, 3.866432, 3.765517, 3.666788, 3.5658894, 3.468703, 3.3619797, 3.2612457, 3.1599743, 3.0651553, 2.9675224, 2.867517, 2.7654264, 2.6686072, 2.567969, 2.4646127, 2.3662403, 2.2672458, 2.1639743, 2.0745115, 1.9656924, 1.8648787, 1.7657936, 1.6727935, 1.5732456, 1.4724212, 1.3685116, 1.2602403, 1.1676978, 1.0685116, 0.97042114, 0.8631499, 0.77142113, 0.6708733, 0.5715966, 0.4670541, 0.36605412, 0.26659665, 0.16896369, 0.065697774, 0.04820052, 0.0, -0.0073742764, 0.030601272, 0.12714916, 0.23242578, 0.33032465, 0.42942578, 0.532697, 0.63269705, 0.7281492, 0.8335109, 0.93724495, 1.0296971, 1.1316066, 1.2371545, 1.3257928, 1.4277024, 1.5306174, 1.6274258, 1.7276067, 1.8318886, 1.9328833, 2.0303407, 2.1277025, 2.2318885, 2.3308885, 2.4322503, 2.535878, 2.6287982, 2.726346, 2.8281653, 2.9279845, 3.0230694, 3.1296172, 3.2239845, 3.3288887, 3.4290748, 3.5245376, 3.6306174, 3.7275321, 3.8287132, 3.927261, 4.0291758, 4.1305375, 4.2238994, 4.3312664, 4.4264417, 4.526713, 4.6318994, 4.724176, 4.8276386, 4.928272, 5.0231757, 5.1239953, 5.223724, 5.323995, 5.424453, 5.525362, 5.6235485, 5.7188196, 5.8196335, 5.926277, 6.01749, 6.1050224, 6.1911025, 6.2721086, 6.350471, 6.4473224, 6.5459604, 6.6483274, 6.7456093, 6.8444285, 6.9463434, 7.0396147, 7.14262, 7.2407055, 7.3428917, 7.438078, 7.544721, 7.6421733, 7.736179, 7.8428063, 7.940365, 8.044456, 8.135737, 8.238105, 8.34528, 8.4401045, 8.535737, 8.635019, 8.740381, 8.841929, 8.935025, 9.034754, 9.136668, 9.237302, 9.332578, 9.434307, 9.53195, 9.640855, 9.736493, 9.832408, 9.930227, 10.039142, 10.131232, 10.231051, 10.330429, 10.432243, 10.529791, 10.63352, 10.733876, 10.828158, 10.927254, 11.023445, 11.128621, 11.228897, 11.324446, 11.423089, 11.521903, 11.629541, 11.722456, 11.822546, 11.922919, 12.019738, 12.121285, 12.221015, 12.31711, 12.422573, 12.522929, 12.618567, 12.724754, 12.81894, 12.915212, 13.016307, 13.118669, 13.216222, 13.316589, 13.4159565, 13.515318, 13.616505, 13.713776, 13.812414, 13.918695, 14.010786, 14.115153, 14.212973, 14.31043, 14.411978, 14.509345, 14.609526, 14.71144, 14.808989, 14.913802, 15.003371, 15.105467, 15.200116, 15.30068, 15.393058, 15.495165, 15.591356, 15.688271, 15.788569, 15.884032, 15.984958, 16.078962, 16.182436, 16.27391, 16.371006, 16.464664, 16.565943, 16.668139, 16.761145, 16.85689, 16.952633, 17.05729, 17.152203, 17.247038, 17.349602, 17.444431, 17.5408, 17.639996, 17.735012, 17.839931, 17.930767, 18.02815, 18.12698, 18.220715, 18.320364, 18.421837, 18.516758, 18.616045, 18.714157, 18.814072, 18.907455, 19.00029, 19.098295, 19.200663, 19.297142, 19.39788, 19.493801, 19.586275, 19.679651, 19.78603, 19.881477, 20.000278, 20.127155, 20.245878, 20.368128, 20.487148, 20.583235, 20.680521, 20.781872, 20.877792, 20.979069, 21.07743, 21.175076, 21.282347, 21.371809, 21.475542, 21.57118, 21.67291, 21.771357, 21.87109, 21.97191, 22.070745, 22.170372, 22.269379, 22.376106, 22.464926, 22.569479, 22.672384, 22.772305, 22.868128, 22.968937, 23.07058, 23.16358, 23.269947, 23.36205, 23.46433, 23.56532, 23.66333, 23.759235, 23.867155, 23.965612, 24.05716, 24.155884, 24.263342, 24.362442, 24.460714, 24.558176, 24.659628, 24.759459, 24.852186, 24.95391, 25.053635, 25.158182, 25.257915, 25.351559, 25.454927, 25.548931, 25.651932, 25.753654, 25.850208, 25.953394, 26.056581, 26.147043, 26.247953, 26.350044, 26.44714, 26.549511, 26.648325, 26.74906, 26.848692, 26.940432, 27.045975, 27.1418, 27.238708, 27.341171, 27.44381, 27.545267, 27.636906, 27.744719, 27.841002, 27.944555, 28.041187, 28.13265, 28.232927, 28.33283, 28.433384, 28.533842, 28.63248, 28.734396, 28.839396, 28.928768, 29.03231, 29.13304, 29.229507, 29.332235, 29.426598, 29.531965, 29.580423, 29.612755, 29.64728, 29.691607, 29.729671, 29.764744, 29.805613, 29.843763, 29.878738, 29.876654, 29.886017, 29.881754, 29.850193, 29.813211, 29.771793, 29.740717, 29.69848, 29.662506, 29.62344, 29.586565, 29.546526, 29.454744, 29.360846, 29.253382, 29.158281, 29.059101, 28.961727, 28.858818, 28.759722, 28.655186, 28.560537, 28.461723, 28.36126, 28.261084, 28.168255, 28.060797, 27.96107, 27.859068, 27.758966, 27.657244, 27.569328, 27.464962, 27.360596, 27.27241, 27.17177, 27.07177, 26.971313, 26.873674, 26.775764, 26.669403, 26.563574, 26.469482, 26.368025, 26.266478, 26.169834, 26.078472, 25.971563, 25.875004, 25.772552, 25.670004, 25.572638, 25.471632, 25.374456, 25.276903, 25.177631, 25.081078, 24.978525, 24.88443, 24.77652, 24.683344, 24.582062, 24.485147, 24.38487, 24.279062, 24.177961, 24.079689, 23.979599, 23.886322, 23.777233, 23.687593, 23.581488, 23.48604, 23.384127, 23.288488, 23.184212, 23.086834, 22.985659, 22.886477, 22.790104, 22.686556, 22.58629, 22.488918, 22.3941, 22.29236, 22.189919, 22.092999, 21.994902, 21.893812, 21.792625, 21.694088, 21.59235, 21.49863, 21.397068, 21.293348, 21.196524, 21.0997, 20.9947, 20.89579, 20.798689, 20.701242, 20.600412, 20.503046, 20.401136, 20.294594, 20.20195, 20.105131, 20.002398, 19.90676, 19.800934, 19.703669, 19.60539, 19.506657, 19.404295, 19.305471, 19.206018, 19.112652, 19.010918, 18.905918, 18.809828, 18.712456, 18.610184, 18.504637, 18.40754, 18.311901, 18.207354, 18.116348, 18.010445, 17.914625, 17.8138, 17.713434, 17.611885, 17.511248, 17.422699, 17.313423, 17.213789, 17.11069, 17.015944, 16.91578, 16.816774, 16.716045, 16.621677, 16.515497, 16.415758, 16.315577, 16.212849, 16.128843, 16.02339, 15.920018, 15.821662, 15.727843, 15.625742, 15.526646, 15.431284, 15.33055, 15.230816, 15.1187315, 15.024918, 14.924635, 14.825279, 14.73154, 14.630268, 14.527444, 14.42462, 14.332257, 14.229896, 14.1328, 14.029524, 13.936518, 13.832422, 13.732518, 13.632332, 13.531241, 13.427423, 13.332422, 13.23305, 13.132045, 13.032492, 12.933316, 12.838768, 12.738491, 12.636034, 12.540029, 12.433215, 12.3370285, 12.238481, 12.139757, 12.0405655, 11.943922, 11.840651, 11.737922, 11.646454, 11.540374, 11.445188, 11.346273, 11.239188, 11.14472, 11.042454, 10.949539, 10.842991, 10.750443, 10.642991, 10.551076, 10.446438, 10.343348, 10.24998, 10.145699, 10.050246, 9.95206, 9.851964, 9.747246, 9.651331, 9.547326, 9.450231, 9.349134, 9.253224, 9.156762, 9.045587, 8.953214, 8.856853, 8.756852, 8.657757, 8.551305, 8.456209, 8.36039, 8.258474, 8.153746, 8.055017, 7.9611025, 7.8589106, 7.760464, 7.659272, 7.566629, 7.4600067, 7.3640914, 7.2653627, 7.159363, 7.0622673, 6.9633574, 6.8609905, 6.7659, 6.6604424, 6.5604424, 6.462889, 6.3714104, 6.295229, 6.200686, 6.117696, 6.0296955, 5.9418387, 5.844105, 5.7434716, 5.6431103, 5.5399294, 5.4409237, 5.342653, 5.2487326, 5.1440144, 5.045913, 4.9441047, 4.8419237, 4.74219, 4.645376, 4.538647, 4.445738, 4.338924, 4.243456, 4.1437325, 4.04428, 3.9461899, 3.843461, 3.7472749, 3.6419187, 3.541376, 3.4438174, 3.3507323, 3.246094, 3.14436, 3.0438175, 2.9421844, 2.8465462, 2.7426312, 2.6437216, 2.543993, 2.440908, 2.342908, 2.2470887, 2.1450887, 2.0428174, 1.9406313, 1.8428972, 1.7461791, 1.648812, 1.5405354, 1.4445407, 1.3389078, 1.2465354, 1.1488013, 1.0432642, 0.9482588, 0.84608334, 0.7458971, 0.6426205, 0.55153006, 0.4522642, 0.3461684, 0.24598756, 0.14471094, 0.047897134, 0.0, -0.0019061053, 0.095024884, 0.19575362, 0.291126, 0.39557812, 0.49710995, 0.59466857, 0.6970249, 0.8008387, 0.8955728, 0.9942111, 1.0963919, 1.198759, 1.297211, 1.3996578, 1.5030249, 1.5945781, 1.6984878, 1.7965728, 1.8925781, 1.9984823, 2.0946686, 2.1912217, 2.2974877, 2.3968654, 2.4936686, 2.5925834, 2.6943972, 2.7982163, 2.8970356, 2.9943123, 3.090493, 3.1961315, 3.288142, 3.3919559, 3.4926794, 3.595041, 3.6942217, 3.7966793, 3.8841367, 3.9926846, 4.097142, 4.1918654, 4.298147, 4.392413, 4.492679, 4.5895944, 4.693052, 4.793605, 4.8885994, 4.99369, 5.085323, 5.1956954, 5.289786, 5.400238, 5.488605, 5.5939612, 5.694062, 5.7859664, 5.8876104, 5.988791, 6.0848813, 6.194961, 6.2956104, 6.3898764, 6.491062, 6.588153, 6.6898813, 6.7858815, 6.8817964, 6.989791, 7.08961, 7.1892486, 7.2896104, 7.39152, 7.4863443, 7.5838923, 7.6912484, 7.7840676, 7.885525, 7.9843497, 8.086616, 8.18635, 8.28626, 8.389259, 8.483073, 8.589344, 8.679078, 8.787079, 8.886988, 8.989615, 9.08435, 9.187807, 9.285185, 9.384536, 9.477637, 9.584531, 9.6809025, 9.7901745, 9.882445, 9.98918, 10.0898075, 10.184004, 10.28027, 10.3851795, 10.486456, 10.587542, 10.6851845, 10.782913, 10.8915415, 10.986637, 11.083095, 11.19018, 11.284642, 11.384371, 11.487547, 11.581914, 11.688637, 11.7900095, 11.8837385, 11.98619, 12.081828, 12.184738, 12.276105, 12.383648, 12.481105, 12.589733, 12.682738, 12.783105, 12.880743, 12.986653, 13.077467, 13.180472, 13.28402, 13.377292, 13.48202, 13.582387, 13.679839, 13.782929, 13.88093, 13.980749, 14.082568, 14.177658, 14.274116, 14.376574, 14.486472, 14.577749, 14.6827545, 14.779935, 14.877308, 14.977212, 15.079211, 15.1835785, 15.272398, 15.38094, 15.475398, 15.571307, 15.678584, 15.774307, 15.877042, 15.978222, 16.077951, 16.178583, 16.278765, 16.379223, 16.471685, 16.577589, 16.684313, 16.77659, 16.878319, 16.974686, 17.071775, 17.175589, 17.275408, 17.375685, 17.479408, 17.576595, 17.673046, 17.773499, 17.869686, 17.97369, 18.07678, 18.177324, 18.271152, 18.378696, 18.473877, 18.57669, 18.674702, 18.774696, 18.87161, 18.972254, 19.0757, 19.161615, 19.27461, 19.37407, 19.471893, 19.571249, 19.67143, 19.772615, 19.874792, 19.973797, 20.074339, 20.172525, 20.269163, 20.369255, 20.464165, 20.566711, 20.667892, 20.77135, 20.869532, 20.971079, 21.066084, 21.168808, 21.268452, 21.367899, 21.472988, 21.56718, 21.663265, 21.762457, 21.86817, 21.964903, 22.065903, 22.167265, 22.27136, 22.371628, 22.466, 22.567722, 22.669096, 22.767372, 22.868366, 22.963186, 23.068457, 23.167913, 23.271282, 23.365818, 23.468372, 23.56683, 23.66265, 23.76665, 23.8651, 23.967106, 24.06283, 24.17028, 24.267015, 24.358738, 24.460297, 24.562382, 24.664473, 24.761484, 24.860388, 24.963026, 25.061659, 25.165388, 25.263025, 25.360207, 25.457394, 25.553392, 25.666117, 25.761936, 25.861488, 25.96276, 26.05277, 26.16158, 26.265303, 26.367212, 26.464941, 26.560038, 26.664404, 26.760307, 26.850319, 26.95877, 27.05559, 27.15859, 27.255962, 27.354319, 27.458319, 27.555138, 27.656048, 27.756052, 27.855234, 27.960415, 28.060862, 28.148245, 28.255144, 28.36324, 28.46142, 28.557867, 28.647335, 28.754877, 28.859781, 28.956244, 29.057516, 29.157068, 29.254515, 29.357334, 29.456882, 29.548367, 29.58913, 29.635105, 29.669527, 29.713678, 29.740208, 29.777353, 29.825233, 29.853926, 29.89336, 29.933605, 29.969847, 30.003813, 30.051693, 30.046703, 30.026178, 29.98613, 29.952238, 29.905907, 29.869383, 29.833961, 29.80017, 29.757298, 29.726046, 29.681889, 29.647652, 29.616219, 29.570532, 29.499014, 29.38911, 29.297377, 29.199743, 29.102652, 28.997375, 28.899828, 28.801376, 28.69628, 28.603008, 28.497828, 28.399733, 28.301281, 28.201456, 28.098185, 27.996733, 27.900461, 27.799913, 27.69845, 27.599552, 27.498371, 27.402908, 27.30309, 27.205093, 27.10136, 27.001625, 26.90627, 26.803806, 26.700626, 26.60453, 26.500355, 26.404625, 26.305445, 26.20262, 26.106802, 26.007439, 25.902983, 25.803982, 25.701439, 25.604078, 25.498169, 25.402163, 25.300259, 25.20044, 25.103615, 24.999079, 24.90643, 24.802887, 24.70752, 24.607332, 24.508429, 24.405882, 24.304338, 24.209509, 24.105423, 24.008419, 23.907423, 23.804695, 23.703876, 23.603056, 23.504593, 23.40778, 23.304508, 23.2086, 23.103418, 23.004955, 22.912413, 22.80705, 22.710594, 22.60396, 22.510962, 22.406775, 22.309227, 22.207148, 22.111317, 22.00886, 21.916216, 21.806046, 21.709679, 21.609493, 21.506311, 21.410397, 21.316584, 21.210407, 21.111403, 21.014307, 20.912577, 20.812035, 20.704493, 20.61802, 20.51712, 20.40703, 20.313215, 20.216206, 20.114843, 20.016838, 19.909391, 19.810572, 19.717567, 19.615385, 19.517656, 19.410662, 19.31102, 19.218296, 19.112747, 19.012562, 18.917662, 18.817741, 18.713743, 18.614477, 18.515461, 18.41547, 18.314291, 18.215923, 18.1181, 18.015928, 17.918652, 17.818913, 17.714924, 17.616827, 17.510279, 17.41855, 17.316456, 17.211552, 17.120092, 17.018188, 16.91746, 16.819094, 16.710646, 16.615004, 16.518093, 16.423178, 16.32028, 16.215454, 16.125816, 16.020636, 15.918449, 15.815992, 15.72145, 15.623088, 15.515992, 15.422626, 15.315721, 15.219535, 15.120263, 15.022907, 14.918088, 14.823896, 14.723716, 14.6195345, 14.51954, 14.419349, 14.325801, 14.211896, 14.117529, 14.023077, 13.9174385, 13.810801, 13.721615, 13.625886, 13.518615, 13.422609, 13.323439, 13.218518, 13.121519, 13.020705, 12.923699, 12.823061, 12.718615, 12.624248, 12.523248, 12.420694, 12.324332, 12.221795, 12.124237, 12.025327, 11.923699, 11.818056, 11.72605, 11.623423, 11.525322, 11.420513, 11.325236, 11.22496, 11.129056, 11.02505, 10.928604, 10.8230505, 10.729231, 10.62496, 10.527141, 10.422875, 10.328321, 10.226859, 10.125141, 10.02704, 9.927407, 9.825046, 9.728221, 9.623774, 9.53322, 9.422401, 9.32704, 9.227582, 9.128402, 9.024864, 8.9269495, 8.828407, 8.72513, 8.628854, 8.529582, 8.427763, 8.329311, 8.230667, 8.122673, 8.034848, 7.9286675, 7.8259387, 7.726029, 7.630215, 7.528582, 7.429481, 7.329391, 7.234566, 7.127125, 7.0301194, 6.9287524, 6.831029, 6.726481, 6.6350236, 6.5322046, 6.4327526, 6.334476, 6.234205, 6.1271195, 6.0257473, 5.927933, 5.8331194, 5.7291994, 5.630109, 5.5321994, 5.4285665, 5.3330183, 5.232199, 5.1352897, 5.0315557, 4.9280186, 4.830832, 4.7351036, 4.636832, 4.5363746, 4.4321938, 4.3350024, 4.2339067, 4.1352787, 4.036098, 3.9280982, 3.8305502, 3.733731, 3.6310024, 3.5319173, 3.4330022, 3.3320076, 3.2330928, 3.1330926, 3.0375395, 2.935545, 2.8349066, 2.7326353, 2.6330023, 2.5358162, 2.4309118, 2.3354545, 2.2402735, 2.138183, 2.0350873, 1.9300821, 1.8381778, 1.7360767, 1.6379863, 1.5387204, 1.4376299, 1.3368107, 1.2344544, 1.1327204, 1.0407096, 0.9372629, 0.84053415, 0.7378054, 0.63734794, 0.53889585, 0.43589583, 0.33661386, 0.23925216, 0.13834794, 0.03925217, 0.07309346, 0.0, 0.083452694, 0.16571918, 0.25942174, 0.35988456, 0.45715582, 0.5533367, 0.65179414, 0.7557995, 0.8557995, 0.9590761, 1.049624, 1.1492623, 1.2585282, 1.3554431, 1.4565336, 1.5554485, 1.6531719, 1.7577251, 1.8471029, 1.9481933, 2.0483634, 2.1514592, 2.2501879, 2.351922, 2.4453743, 2.5512836, 2.6494646, 2.746289, 2.8515604, 2.9439328, 3.04847, 3.1458316, 3.2414806, 3.3519328, 3.4495764, 3.5410285, 3.6472094, 3.7482998, 3.8433955, 3.9436774, 4.045582, 4.1399436, 4.24322, 4.3458586, 4.441592, 4.543864, 4.647401, 4.744146, 4.842502, 4.9444118, 5.0338798, 5.1379647, 5.2356086, 5.338061, 5.4383373, 5.5353374, 5.638795, 5.7356086, 5.8369756, 5.937981, 6.0341616, 6.1412573, 6.2389865, 6.3430715, 6.4365287, 6.5419865, 6.6379914, 6.7354436, 6.8391776, 6.9297204, 7.0343585, 7.1263695, 7.2374597, 7.331651, 7.434731, 7.531375, 7.630923, 7.738098, 7.8300185, 7.9313803, 8.030933, 8.131114, 8.234481, 8.328119, 8.431024, 8.526672, 8.631758, 8.725035, 8.827667, 8.919683, 9.018248, 9.121806, 9.217269, 9.31637, 9.414747, 9.510306, 9.607136, 9.706966, 9.800982, 9.897535, 10.001009, 10.094839, 10.190121, 10.300594, 10.3887005, 10.490344, 10.585994, 10.68518, 10.781829, 10.877127, 10.974408, 11.070058, 11.16852, 11.262712, 11.366728, 11.467739, 11.563207, 11.654494, 11.750143, 11.848431, 11.950627, 12.048271, 12.151463, 12.250755, 12.346394, 12.439601, 12.542069, 12.633989, 12.732904, 12.830197, 12.933118, 13.024586, 13.121596, 13.211698, 13.317352, 13.419182, 13.516102, 13.606661, 13.713214, 13.829006, 13.961627, 14.071973, 14.188137, 14.308497, 14.408413, 14.508237, 14.605328, 14.707966, 14.8024235, 14.909424, 15.005333, 15.105344, 15.20344, 15.305796, 15.409349, 15.50562, 15.596902, 15.698812, 15.800993, 15.89836, 16.001455, 16.099737, 16.198462, 16.300642, 16.3991, 16.493738, 16.602375, 16.69811, 16.79393, 16.893116, 16.991663, 17.092579, 17.19012, 17.293125, 17.397217, 17.494318, 17.595493, 17.6925, 17.794228, 17.886509, 17.987051, 18.09842, 18.19051, 18.287971, 18.38688, 18.489424, 18.588882, 18.688435, 18.781893, 18.88217, 18.987898, 19.086718, 19.183989, 19.281004, 19.381819, 19.48609, 19.577732, 19.68428, 19.777287, 19.87683, 19.979744, 20.07693, 20.181381, 20.281473, 20.374302, 20.48212, 20.577387, 20.677307, 20.77567, 20.872505, 20.980047, 21.07386, 21.174137, 21.277596, 21.371956, 21.47242, 21.57733, 21.676243, 21.766605, 21.87043, 21.967978, 22.06843, 22.166712, 22.265717, 22.371254, 22.4649, 22.567356, 22.66309, 22.76436, 22.866638, 22.964367, 23.071089, 23.163378, 23.26293, 23.362473, 23.41364, 23.458332, 23.488037, 23.529001, 23.561983, 23.608496, 23.640562, 23.678255, 23.718779, 23.758924, 23.794804, 23.832603, 23.868383, 23.904263, 23.903822, 23.884207, 23.843332, 23.811176, 23.771658, 23.740587, 23.696712, 23.65902, 23.620314, 23.583616, 23.549011, 23.503675, 23.46971, 23.430458, 23.401499, 23.306791, 23.199966, 23.106419, 23.005865, 22.906408, 22.806316, 22.71022, 22.610493, 22.517035, 22.413307, 22.312939, 22.21003, 22.109663, 22.014296, 21.917658, 21.814291, 21.711552, 21.614832, 21.5101, 21.417912, 21.317455, 21.216726, 21.124992, 21.015636, 20.920986, 20.821167, 20.724716, 20.622173, 20.5228, 20.42244, 20.320343, 20.219614, 20.12488, 20.021881, 19.925327, 19.824965, 19.722424, 19.627954, 19.529316, 19.42704, 19.323046, 19.228312, 19.12322, 19.027029, 18.930487, 18.829662, 18.72857, 18.635662, 18.534746, 18.427475, 18.337831, 18.236109, 18.131645, 18.032555, 17.932913, 17.836365, 17.736273, 17.636635, 17.5379, 17.4349, 17.334263, 17.237896, 17.13698, 17.039986, 16.9368, 16.836885, 16.741789, 16.641975, 16.54397, 16.442965, 16.339874, 16.244501, 16.141863, 16.041502, 15.944316, 15.84413, 15.742125, 15.641406, 15.542582, 15.445577, 15.346666, 15.2513, 15.148028, 15.042113, 14.947475, 14.844204, 14.75038, 14.646103, 14.552007, 14.448555, 14.348374, 14.249273, 14.151448, 14.053459, 13.952821, 13.84872, 13.755268, 13.65463, 13.550896, 13.452714, 13.351619, 13.255884, 13.15507, 13.055432, 12.95806, 12.852698, 12.7516985, 12.656151, 12.555969, 12.454592, 12.358235, 12.253321, 12.156682, 12.058321, 11.964858, 11.859868, 11.760677, 11.661502, 11.561768, 11.456948, 11.363581, 11.263395, 11.162943, 11.059853, 10.964028, 10.866841, 10.766395, 10.661203, 10.565294, 10.460566, 10.363023, 10.268289, 10.16656, 10.072373, 9.963736, 9.864012, 9.769283, 9.669368, 9.566187, 9.471002, 9.370549, 9.268809, 9.173001, 9.0713625, 8.968086, 8.868905, 8.773442, 8.673799, 8.567815, 8.467533, 8.371076, 8.273985, 8.173613, 8.073613, 7.974437, 7.872698, 7.779788, 7.6704264, 7.5748787, 7.476698, 7.3732347, 7.26932, 7.1734157, 7.0795064, 6.9715915, 6.8783145, 6.776134, 6.6738625, 6.572134, 6.4785857, 6.37749, 6.2775807, 6.1834903, 6.083666, 5.9765754, 5.8832135, 5.7833943, 5.679389, 5.580389, 5.4927454, 5.383745, 5.284745, 5.1871123, 5.084011, 4.9824634, 4.8801866, 4.782192, 4.682373, 4.5847454, 4.4827294, 4.383639, 4.284543, 4.184729, 4.0849953, 3.9844472, 3.8886335, 3.7936227, 3.6858144, 3.592894, 3.4858036, 3.386623, 3.2881653, 3.1918888, 3.0879738, 2.9864366, 2.8880696, 2.7887876, 2.6963408, 2.5933301, 2.4894207, 2.3879738, 2.2894206, 2.1929631, 2.095692, 1.996229, 1.8836865, 1.7925056, 1.6944045, 1.5946811, 1.4942291, 1.3881279, 1.2856811, 1.1945853, 1.0931278, 0.99067044, 0.89303213, 0.79385126, 0.69121295, 0.59530336, 0.49666506, 0.39411184, 0.3017448, 0.20380844, 0.1157228, 0.03546166, 0.0, 0.037996963, 0.13307668, 0.23272035, 0.3341778, 0.42781612, 0.5339065, 0.6315448, 0.7278161, 0.8326353, 0.9341778, 1.0330874, 1.1304544, 1.233731, 1.3274544, 1.435731, 1.5306406, 1.6318269, 1.7336407, 1.8305502, 1.9348161, 2.0311832, 2.1330926, 2.2279172, 2.3318214, 2.431731, 2.5339227, 2.629465, 2.7294652, 2.8313801, 2.9314597, 3.028194, 3.1283748, 3.2288322, 3.331013, 3.4292045, 3.5252895, 3.6305609, 3.7300076, 3.8322897, 3.93138, 4.0281034, 4.1306567, 4.228662, 4.3276567, 4.4312897, 4.5312896, 4.630832, 4.7334704, 4.825662, 4.93038, 5.0265718, 5.132024, 5.2298427, 5.328843, 5.4297576, 5.528295, 5.6265717, 5.7237525, 5.8278484, 5.9314814, 6.021327, 6.1103225, 6.1931367, 6.2733183, 6.3580475, 6.4526277, 6.5459943, 6.6498985, 6.75, 6.8492713, 6.945824, 7.045367, 7.150372, 7.2458353, 7.342197, 7.4447393, 7.5446544, 7.644931, 7.7457447, 7.843388, 7.9403033, 8.043122, 8.138123, 8.237213, 8.343128, 8.4394045, 8.542862, 8.642314, 8.738404, 8.843777, 8.934235, 9.03724, 9.13533, 9.2363405, 9.332606, 9.442698, 9.538516, 9.64134, 9.735075, 9.838803, 9.93116, 10.032166, 10.135984, 10.239995, 10.327447, 10.435081, 10.532182, 10.634362, 10.731554, 10.8320055, 10.9240055, 11.030368, 11.13074, 11.225192, 11.327106, 11.434745, 11.533559, 11.624479, 11.725118, 11.826846, 11.929575, 12.028298, 12.124857, 12.224495, 12.319676, 12.430405, 12.52441, 12.619586, 12.722873, 12.821059, 12.920144, 13.017969, 13.120511, 13.2239685, 13.322427, 13.419703, 13.512346, 13.620166, 13.713352, 13.813714, 13.91199, 14.017171, 14.1141815, 14.217814, 14.316086, 14.413826, 14.511644, 14.612639, 14.7149105, 14.808379, 14.914741, 15.009576, 15.113405, 15.209597, 15.3015175, 15.403906, 15.5058155, 15.591741, 15.692938, 15.788406, 15.889321, 15.985342, 16.08054, 16.182455, 16.278475, 16.376396, 16.468954, 16.567146, 16.661806, 16.762997, 16.862913, 16.959652, 17.059679, 17.153412, 17.257061, 17.350986, 17.447727, 17.546919, 17.648115, 17.744036, 17.836046, 17.9347, 18.033627, 18.130722, 18.233286, 18.329659, 18.419222, 18.521967, 18.617887, 18.71236, 18.811626, 18.90793, 19.00967, 19.107409, 19.198143, 19.301435, 19.39826, 19.490648, 19.593473, 19.686043, 19.791138, 19.885857, 20.006653, 20.122818, 20.252163, 20.373875, 20.489891, 20.586252, 20.683996, 20.78281, 20.885258, 20.975716, 21.080545, 21.185453, 21.280464, 21.381002, 21.476284, 21.578375, 21.676657, 21.776114, 21.874475, 21.978386, 22.070572, 22.176752, 22.27812, 22.375305, 22.477486, 22.570763, 22.677221, 22.778955, 22.875046, 22.974949, 23.070417, 23.170326, 23.270603, 23.37152, 23.466608, 23.564892, 23.672434, 23.765987, 23.864353, 23.967264, 24.065722, 24.166264, 24.265455, 24.36473, 24.462912, 24.56846, 24.656828, 24.760923, 24.863098, 24.96193, 25.062561, 25.161295, 25.2563, 25.353115, 25.457222, 25.559584, 25.661488, 25.759407, 25.855774, 25.952322, 26.052694, 26.15496, 26.250328, 26.36087, 26.448242, 26.54979, 26.652977, 26.752802, 26.852348, 26.947168, 27.052536, 27.149174, 27.243992, 27.352907, 27.451275, 27.550184, 27.638945, 27.675644, 27.719242, 27.755222, 27.791012, 27.829157, 27.867313, 27.907646, 27.943617, 27.982592, 28.01929, 28.058798, 28.057707, 28.029758, 27.99732, 27.966429, 27.922651, 27.88577, 27.839258, 27.808655, 27.7725, 27.733704, 27.689474, 27.655226, 27.590326, 27.488226, 27.388859, 27.282774, 27.193577, 27.092396, 26.986034, 26.889023, 26.793928, 26.698109, 26.593842, 26.496464, 26.391554, 26.297188, 26.197464, 26.095093, 25.998905, 25.893543, 25.792543, 25.69799, 25.59672, 25.500448, 25.40516, 25.302252, 25.203161, 25.101522, 25.001251, 24.901884, 24.801054, 24.70106, 24.602144, 24.501144, 24.408676, 24.303959, 24.212309, 24.109762, 24.013304, 23.905937, 23.814486, 23.706757, 23.612938, 23.514927, 23.412378, 23.315464, 23.21147, 23.110464, 23.01282, 22.910181, 22.82464, 22.717724, 22.613544, 22.512358, 22.411533, 22.316538, 22.214613, 22.123346, 22.025166, 21.921787, 21.81825, 21.716156, 21.62197, 21.521053, 21.424597, 21.317055, 21.22241, 21.118044, 21.026587, 20.924671, 20.824219, 20.72376, 20.627762, 20.526028, 20.436117, 20.326756, 20.226847, 20.132654, 20.027836, 19.931198, 19.827559, 19.733187, 19.631283, 19.527735, 19.435368, 19.331001, 19.230724, 19.133537, 19.035719, 18.940893, 18.837803, 18.736065, 18.633888, 18.535526, 18.434889, 18.340696, 18.240788, 18.134783, 18.035877, 17.937963, 17.838415, 17.74159, 17.641048, 17.53732, 17.437134, 17.345495, 17.239952, 17.140394, 17.04685, 16.93957, 16.847027, 16.750378, 16.646835, 16.544655, 16.441744, 16.349281, 16.24801, 16.1441, 16.045366, 15.951362, 15.849723, 15.751628, 15.649367, 15.553808, 15.448627, 15.351984, 15.244074, 15.152436, 15.054069, 14.95525, 14.854797, 14.753244, 14.65851, 14.558148, 14.456691, 14.36168, 14.255329, 14.153409, 14.053776, 13.954957, 13.857771, 13.759584, 13.65558, 13.562765, 13.457212, 13.362117, 13.263569, 13.163744, 13.063287, 12.964382, 12.862105, 12.767197, 12.667281, 12.56518, 12.466643, 12.368366, 12.2665415, 12.165999, 12.069361, 11.971898, 11.869984, 11.77026, 11.665723, 11.570797, 11.4692545, 11.362701, 11.266616, 11.172882, 11.074972, 10.970329, 10.875787, 10.771329, 10.6746, 10.573595, 10.4749565, 10.377132, 10.273228, 10.172674, 10.077403, 9.976132, 9.877573, 9.777297, 9.676387, 9.575393, 9.482658, 9.380653, 9.280925, 9.172563, 9.087924, 8.980552, 8.880648, 8.782547, 8.682365, 8.582281, 8.486908, 8.385823, 8.288175, 8.18544, 8.08535, 7.9855304, 7.8857965, 7.79235, 7.6878815, 7.585621, 7.4904346, 7.3875146, 7.2886047, 7.1923285, 7.0907855, 6.9865146, 6.891413, 6.796408, 6.6914983, 6.5946794, 6.4974027, 6.3933015, 6.315487, 6.226141, 6.14205, 6.054778, 5.9646287, 5.8663573, 5.772081, 5.671985, 5.569538, 5.4683523, 5.367533, 5.276352, 5.1669903, 5.068246, 4.9717083, 4.8698893, 4.770267, 4.675347, 4.570799, 4.4718785, 4.371884, 4.2740703, 4.168884, 4.076698, 3.9657085, 3.8716073, 3.773251, 3.6734264, 3.5749743, 3.4717085, 3.3747828, 3.2696073, 3.1676128, 3.0739799, 2.9713306, 2.8690596, 2.7706978, 2.678884, 2.5810647, 2.4696126, 2.373235, 2.272602, 2.1736073, 2.0679636, 1.9708786, 1.8706924, 1.7746924, 1.6759636, 1.577687, 1.4763147, 1.3761499, 1.276602, 1.1744158, 1.0795009, 0.9741445, 0.8736871, 0.7712296, 0.6722296, 0.57158595, 0.47431466, 0.37786257, 0.2757775, 0.17413382, 0.077947624, 0.11206018, 0.0, -0.0010125868, 0.08569531, 0.18788151, 0.28269532, 0.3746156, 0.48424855, 0.579424, 0.67707306, 0.7752432, 0.8806102, 0.9786156, 1.0822539, 1.1731635, 1.279339, 1.3813443, 1.4796156, 1.5762432, 1.683988, 1.7819773, 1.8825198, 1.9756103, 2.0773497, 2.176706, 2.2736208, 2.377706, 2.4818017, 2.5773497, 2.6754456, 2.7786317, 2.8818018, 2.9716318, 3.0798018, 3.171988, 3.2795358, 3.3770838, 3.4759934, 3.5737221, 3.6729083, 3.7785358, 3.8789933, 3.982621, 4.078089, 4.179807, 4.277174, 4.382536, 4.474632, 4.576451, 4.674451, 4.772547, 4.8758125, 4.977722, 5.070914, 5.173993, 5.279185, 5.3786426, 5.476642, 5.5823655, 5.67536, 5.771004, 5.877999, 5.9741797, 6.0581694, 6.1477976, 6.234245, 6.3104315, 6.3988686, 6.5027833, 6.593608, 6.6985226, 6.791065, 6.894608, 6.9939857, 7.0962462, 7.1949854, 7.2953525, 7.3985333, 7.4950867, 7.5995336, 7.693911, 7.787369, 7.8963633, 7.9891825, 8.091996, 8.19073, 8.290464, 8.3893795, 8.48947, 8.589837, 8.690843, 8.786114, 8.886571, 8.986481, 9.082666, 9.183028, 9.287401, 9.38231, 9.485226, 9.578677, 9.680316, 9.782959, 9.87605, 9.983513, 10.0762415, 10.186236, 10.277959, 10.376694, 10.480603, 10.581518, 10.677252, 10.779167, 10.880161, 10.975981, 11.075986, 11.1793585, 11.274173, 11.3708105, 11.477359, 11.572178, 11.674183, 11.771189, 11.87664, 11.967103, 12.0760975, 12.167109, 12.280917, 12.374199, 12.471013, 12.575396, 12.672476, 12.770396, 12.866753, 12.970029, 13.071577, 13.16795, 13.270944, 13.369774, 13.463136, 13.5636835, 13.664875, 13.762231, 13.86297, 13.9672365, 14.062699, 14.161518, 14.264343, 14.35979, 14.457258, 14.562982, 14.652082, 14.761806, 14.862716, 14.955545, 15.051918, 15.154928, 15.248306, 15.3485985, 15.442971, 15.54271, 15.641631, 15.741376, 15.837578, 15.93504, 16.028866, 16.127237, 16.227074, 16.325636, 16.422918, 16.517212, 16.616133, 16.708052, 16.809973, 16.90844, 17.004547, 17.102467, 17.204025, 17.30368, 17.398685, 17.495893, 17.593988, 17.691633, 17.786472, 17.883026, 17.983957, 18.08215, 18.175255, 18.269266, 18.376276, 18.469378, 18.566128, 18.66223, 18.75733, 18.859985, 18.961996, 19.058283, 19.152847, 19.251406, 19.343779, 19.444155, 19.540438, 19.635279, 19.73947, 19.8363, 19.948309, 20.065845, 20.187553, 20.307085, 20.427057, 20.529232, 20.632961, 20.731781, 20.83387, 20.929148, 21.029068, 21.1257, 21.237152, 21.327068, 21.424892, 21.52844, 21.620356, 21.724535, 21.828535, 21.916632, 22.027721, 22.123636, 22.224184, 22.329733, 22.422106, 22.518833, 22.61993, 22.721647, 22.81802, 22.9242, 23.019115, 23.121387, 23.215845, 23.313036, 23.411585, 23.51668, 23.613499, 23.715137, 23.816408, 23.921505, 24.015871, 24.108961, 24.213062, 24.313515, 24.411612, 24.50734, 24.60916, 24.707531, 24.803988, 24.907255, 25.00808, 25.109716, 25.20509, 25.309818, 25.403461, 25.503191, 25.60583, 25.703924, 25.803919, 25.901201, 26.005291, 26.099936, 26.205574, 26.300303, 26.40485, 26.503126, 26.592585, 26.702494, 26.793867, 26.899408, 26.995504, 27.097324, 27.195059, 27.293882, 27.398335, 27.49625, 27.59152, 27.696068, 27.790073, 27.893984, 27.988724, 28.090357, 28.187271, 28.29309, 28.38782, 28.492096, 28.581469, 28.689734, 28.785654, 28.883383, 28.98666, 29.085299, 29.190388, 29.290575, 29.38239, 29.479128, 29.560432, 29.600674, 29.637281, 29.668072, 29.705961, 29.7433, 29.790443, 29.821873, 29.861113, 29.89936, 29.931879, 29.967571, 29.96821, 29.970047, 29.937168, 29.89983, 29.862223, 29.821527, 29.780373, 29.747126, 29.70724, 29.668184, 29.63839, 29.595419, 29.555183, 29.469337, 29.37761, 29.277874, 29.176964, 29.086603, 28.981688, 28.880322, 28.782045, 28.676226, 28.585667, 28.485401, 28.384401, 28.282581, 28.19039, 28.090023, 27.987108, 27.887384, 27.791199, 27.68738, 27.588379, 27.493008, 27.384544, 27.28864, 27.19455, 27.090538, 26.991545, 26.891533, 26.801167, 26.691076, 26.591528, 26.495342, 26.395618, 26.297976, 26.194788, 26.097511, 25.99697, 25.894236, 25.800596, 25.695139, 25.593502, 25.497591, 25.398863, 25.300406, 25.205948, 25.098846, 25.002123, 24.905842, 24.803757, 24.705933, 24.606295, 24.507835, 24.41283, 24.309458, 24.202831, 24.110548, 24.010544, 23.905453, 23.811447, 23.712442, 23.61072, 23.508257, 23.407804, 23.313618, 23.2088, 23.112432, 23.01534, 22.915703, 22.81424, 22.712517, 22.605879, 22.514416, 22.417772, 22.31351, 22.21268, 22.112953, 22.018496, 21.914043, 21.819672, 21.72049, 21.628021, 21.517847, 21.422836, 21.320936, 21.221842, 21.118017, 21.021282, 20.91965, 20.824463, 20.720282, 20.625368, 20.519459, 20.427181, 20.327, 20.224533, 20.124628, 20.026712, 19.930437, 19.822346, 19.723713, 19.630697, 19.528059, 19.432878, 19.336512, 19.233511, 19.135872, 19.027872, 18.93124, 18.835777, 18.731861, 18.637314, 18.533766, 18.432219, 18.33331, 18.237309, 18.135033, 18.03693, 17.935472, 17.836384, 17.73466, 17.634659, 17.535107, 17.438196, 17.338644, 17.243282, 17.137096, 17.042006, 16.939, 16.842632, 16.744898, 16.643446, 16.544447, 16.441526, 16.34808, 16.241802, 16.142984, 16.041431, 15.94834, 15.8447075, 15.748606, 15.645515, 15.557414, 15.445058, 15.349324, 15.248781, 15.1484995, 15.048866, 14.95159, 14.848319, 14.750122, 14.65558, 14.55477, 14.4549465, 14.350845, 14.256845, 14.1561165, 14.056749, 13.958015, 13.859286, 13.754925, 13.651919, 13.551377, 13.459733, 13.355, 13.258361, 13.157361, 13.054356, 12.961084, 12.857441, 12.7552595, 12.658525, 12.56026, 12.463441, 12.367068, 12.263159, 12.166611, 12.063962, 11.962244, 11.862781, 11.766781, 11.669967, 11.565324, 11.4681425, 11.365685, 11.26759, 11.169494, 11.068042, 10.969765, 10.867494, 10.769307, 10.674121, 10.573297, 10.471663, 10.36893, 10.267291, 10.167116, 10.074281, 9.97319, 9.8741, 9.778733, 9.672366, 9.575191, 9.47336, 9.376908, 9.270722, 9.175536, 9.077807, 8.976265, 8.87553, 8.777531, 8.678621, 8.585701, 8.481249, 8.374706, 8.283339, 8.186972, 8.076509, 7.9834185, 7.881328, 7.77861, 7.685046, 7.5896845, 7.481408, 7.3850465, 7.285403, 7.186403, 7.091578, 6.985222, 6.8873014, 6.788482, 6.685291, 6.582211, 6.487477, 6.386014, 6.304375, 6.220758, 6.132491, 6.0573044, 5.9658732, 5.866421, 5.7709637, 5.665421, 5.5667033, 5.465602, 5.3640594, 5.268421, 5.165421, 5.069868, 4.964235, 4.868602, 4.7666817, 4.664235, 4.565687, 4.4657774, 4.3699584, 4.266958, 4.1662297, 4.0714107, 3.9682243, 3.8704104, 3.7674158, 3.6656816, 3.5750487, 3.466687, 3.368405, 3.271134, 3.1679475, 3.0737667, 2.9684105, 2.8650486, 2.776038, 2.6685805, 2.566304, 2.4707615, 2.3713093, 2.275038, 2.1765807, 2.067038, 1.9734901, 1.8695806, 1.7733094, 1.6686656, 1.5706656, 1.4746603, 1.3713039, 1.2659476, 1.1711178, 1.0704795, 0.9755806, 0.8742082, 0.77366567, 0.67211777, 0.57429326, 0.47357523, 0.37058058, 0.26702735, 0.17038903, 0.07320819, 0.03215292];
    F : ARRAY[0..5931] OF REAL := [2.842882, 6.817853, 6.893808, 6.8648725, 6.890191, 6.922743, 6.92636, 6.929977, 6.9516783, 6.915509, 6.890191, 6.9733796, 6.980613, 6.890191, 6.915509, 6.919126, 6.929977, 6.9408274, 6.929977, 6.9480615, 6.991464, 7.020399, 6.9480615, 7.005932, 6.9842305, 6.9986978, 6.991464, 6.9625287, 7.005932, 7.002315, 7.0131655, 6.980613, 7.0131655, 7.0095487, 7.0131655, 6.9733796, 7.0131655, 7.0384836, 7.060185, 7.0457177, 7.096354, 7.092737, 7.0529513, 7.071036, 7.0999713, 7.0638022, 7.1180553, 7.056568, 7.1289062, 7.143374, 7.1180553, 7.1252894, 7.172309, 7.1252894, 7.1614585, 7.0891204, 7.0999713, 7.146991, 7.2229457, 7.1180553, 7.157841, 7.1903934, 7.7654805, 8.412905, 9.027778, 9.707755, 10.304543, 10.250289, 10.235822, 10.250289, 10.304543, 10.279224, 10.358796, 10.297309, 10.420283, 10.4347515, 10.373264, 10.452836, 10.456452, 10.427517, 10.463686, 10.4817705, 10.503472, 10.521557, 10.546875, 10.583044, 10.579427, 10.619213, 10.6119795, 10.644531, 10.666233, 10.734954, 10.734954, 10.698785, 10.774739, 10.78559, 10.807292, 10.778357, 10.756655, 10.821759, 10.850695, 10.807292, 10.847077, 10.904948, 10.8723955, 10.876013, 10.944734, 10.944734, 11.009838, 11.006221, 11.020689, 11.064092, 11.035156, 11.08941, 11.118345, 11.172599, 11.158131, 11.158131, 11.125579, 11.161748, 11.2630205, 11.205151, 11.29919, 11.288339, 11.219618, 11.31004, 11.306423, 11.317274, 11.349827, 11.364294, 11.378761, 11.429399, 11.447483, 11.400463, 11.454717, 11.46195, 11.490886, 11.527055, 11.548756, 11.570457, 11.624711, 11.534288, 11.682581, 11.621094, 11.599392, 11.657263, 11.747685, 11.722367, 11.76577, 11.725984, 11.71875, 11.754919, 11.801939, 11.921296, 12.008101, 12.145544, 12.286603, 12.358941, 12.398726, 12.543403, 12.641059, 12.760417, 12.814671, 12.941261, 13.057002, 13.122107, 13.208912, 13.335504, 13.440393, 13.53805, 13.599537, 13.708044, 13.791233, 13.939526, 14.022714, 14.123987, 14.210793, 14.322917, 14.391638, 14.47121, 14.579717, 14.735243, 14.728009, 14.919704, 14.999276, 15.140336, 15.223524, 15.332031, 15.4296875, 15.530961, 15.625, 15.675636, 15.838397, 15.878182, 15.921586, 16.084347, 16.24349, 16.323061, 16.44242, 16.540075, 16.543692, 16.731771, 16.818577, 16.171152, 15.386285, 14.47121, 13.729745, 12.999132, 12.890625, 12.879774, 12.97743, 12.959346, 12.959346, 13.006366, 12.999132, 13.035301, 13.006366, 13.057002, 13.075087, 13.132957, 13.132957, 13.190827, 13.198061, 13.154658, 13.266783, 13.23423, 13.28125, 13.295717, 13.299335, 13.302952, 13.317419, 13.382524, 13.349971, 13.404224, 13.483796, 13.38614, 13.505498, 13.48018, 13.530816, 13.530816, 13.581452, 13.588686, 13.6067705, 13.632089, 13.635706, 13.661024, 13.726129, 13.711661, 13.722511, 13.726129, 13.776765, 13.740596, 13.838252, 13.831018, 13.838252, 13.906974, 13.935908, 13.932292, 13.939526, 13.986546, 13.964844, 13.993779, 14.1276045, 14.019097, 14.134838, 14.134838, 14.12037, 14.138454, 14.1276045, 14.189092, 14.254195, 14.210793, 14.210793, 14.2578125, 14.290364, 14.290364, 14.348235, 14.326533, 14.395255, 14.431423, 14.420573, 14.413339, 14.478443, 14.521846, 14.507379, 14.576099, 14.514612, 14.572483, 14.58695, 14.561632, 14.699074, 14.662905, 14.69184, 14.742476, 14.767796, 14.800347, 14.78588, 14.850984, 14.803964, 16.030092, 18.514902, 21.050346, 23.488136, 25.99103, 28.47584, 30.9932, 33.449074, 35.92303, 38.465714, 40.93967, 40.990307, 37.807438, 35.337093, 32.7908, 30.35301, 27.846498, 25.343605, 22.887732, 20.330584, 17.896412, 15.379051, 13.136574, 13.111256, 13.049768, 13.111256, 13.049768, 13.0027485, 12.973814, 12.97743, 12.86169, 12.934028, 12.890625, 12.876158, 12.876158, 12.814671, 12.839989, 12.785735, 12.774884, 12.706163, 12.760417, 12.706163, 12.666377, 12.6953125, 12.644676, 12.622974, 12.597656, 12.554254, 12.590423, 12.528935, 12.503617, 12.532552, 12.510851, 12.413195, 12.420428, 12.398726, 12.402344, 12.337239, 12.351707, 12.333623, 12.261285, 12.239583, 12.257668, 12.207031, 12.203414, 12.185329, 12.163629, 12.192564, 12.141927, 12.131077, 12.047888, 12.09129, 12.040654, 12.037037, 11.982783, 12.015336, 11.961082, 11.935764, 11.92853, 11.91768, 11.856193, 11.888744, 11.867043, 11.794704, 11.801939, 11.805555, 11.762153, 11.71875, 11.700665, 11.67173, 11.697048, 11.617476, 11.584925, 11.635561, 11.599392, 11.570457, 11.555989, 11.545139, 11.516204, 11.476418, 11.498119, 11.469184, 11.46195, 11.407697, 11.342592, 11.443866, 11.349827, 11.328125, 11.281105, 11.230469, 11.306423, 11.223235, 11.201533, 11.226851, 11.129195, 11.082176, 11.111111, 11.121962, 11.078559, 11.0496235, 11.082176, 11.006221, 11.103877, 11.038774, 10.99537, 10.933883, 10.966435, 10.915798, 10.89048, 10.854311, 10.923033, 10.814526, 10.8723955, 10.767506, 10.807292, 10.796441, 10.756655, 10.713252, 10.724103, 10.655382, 10.673467, 10.6119795, 10.666233, 10.626447, 10.554109, 10.543258, 10.507089, 10.525173, 10.489005, 10.56496, 10.507089, 10.478154, 10.420283, 10.398582, 10.398582, 10.362413, 10.369647, 10.311776, 10.347945, 10.282842, 10.297309, 10.206886, 10.275608, 10.224971, 10.243055, 10.206886, 10.127315, 10.159867, 10.134548, 10.116464, 10.123698, 10.05136, 10.127315, 10.047743, 10.040509, 10.007957, 10.018807, 10.015191, 9.888599, 9.975405, 9.910301, 9.942853, 9.895833, 9.942853, 9.859664, 9.809028, 9.812645, 9.827112, 9.758391, 9.751158, 9.769242, 9.711371, 9.689671, 9.664351, 9.686053, 9.595631, 9.617332, 9.58478, 9.57393, 9.624566, 9.5703125, 9.505208, 9.4871235, 9.490741, 9.47989, 9.469039, 9.436487, 9.393085, 9.393085, 9.385851, 9.367766, 9.324364, 9.32798, 9.313513, 9.277344, 9.288195, 9.266493, 9.255642, 9.201389, 9.201389, 9.197772, 9.215857, 9.150752, 9.150752, 9.16522, 9.161603, 9.100116, 9.085649, 8.995226, 9.016927, 9.020544, 8.984375, 8.991609, 8.96629, 8.937355, 8.95544, 8.904803, 8.89757, 8.868634, 8.901186, 8.810764, 8.79268, 8.785445, 8.832465, 8.807147, 8.709491, 8.7058735, 8.723958, 8.69864, 8.676939, 8.687789, 8.637153, 8.586516, 8.669704, 8.65162, 8.311632, 7.671441, 7.060185, 6.4127603, 5.754485, 5.5266204, 5.519387, 5.541088, 5.5266204, 5.5483217, 5.46875, 5.4904513, 5.5013022, 5.4868345, 5.494068, 5.4253473, 5.4217305, 5.479601, 5.4868345, 5.396412, 5.4253473, 5.4361978, 5.428964, 5.465133, 5.4217305, 5.432581, 5.4361978, 5.443432, 5.3855615, 5.4217305, 5.4253473, 5.432581, 5.432581, 5.3855615, 5.360243, 5.4000287, 5.3493924, 5.3385415, 5.3385415, 5.331308, 5.342159, 5.342159, 5.4108796, 5.3132234, 5.360243, 5.2987556, 5.327691, 5.3023725, 5.3023725, 5.31684, 5.31684, 5.367477, 5.280671, 5.31684, 5.2842884, 5.291522, 5.255353, 5.331308, 5.2408853, 5.3132234, 5.2842884, 5.230035, 5.2842884, 5.2336516, 5.2336516, -0.014467592, 5.295139, 7.096354, 7.0493345, 7.0782695, 7.060185, 7.0240164, 7.0999713, 7.1180553, 7.0891204, 7.060185, 7.103588, 7.13614, 7.0855036, 7.1289062, 7.1252894, 7.071036, 7.1216726, 7.1903934, 7.107205, 7.1903934, 7.146991, 7.1289062, 7.146991, 7.18316, 7.1867766, 7.1650753, 7.1903934, 7.1976275, 7.18316, 7.168692, 7.2265625, 7.18316, 7.1903934, 7.212095, 7.219329, 7.208478, 7.2229457, 7.2301793, 7.1976275, 7.2554975, 7.244647, 7.2663484, 7.269965, 7.295284, 7.2229457, 7.3350697, 7.2916665, 7.284433, 7.284433, 7.2229457, 7.306134, 7.2989006, 7.280816, 7.8993053, 8.622685, 9.186921, 9.874132, 10.438368, 10.36603, 10.380498, 10.409432, 10.441985, 10.536024, 10.550492, 10.521557, 10.521557, 10.521557, 10.597511, 10.525173, 10.630064, 10.651765, 10.640914, 10.666233, 10.698785, 10.753038, 10.78559, 10.6589985, 10.789207, 10.753038, 10.814526, 10.796441, 10.810908, 10.876013, 10.865162, 10.912182, 10.908565, 10.980903, 10.912182, 10.919415, 10.98452, 10.941117, 11.017072, 11.053241, 11.031539, 11.129195, 11.107494, 11.13643, 11.121962, 11.187066, 11.201533, 11.2160015, 11.219618, 11.288339, 11.295573, 11.244936, 11.266638, 11.338976, 11.364294, 11.302807, 11.378761, 11.407697, 11.396846, 11.433015, 11.454717, 11.480035, 11.476418, 11.501736, 11.51982, 11.505353, 11.548756, 11.588542, 11.599392, 11.6066265, 11.631945, 11.610243, 11.733217, 11.71875, 11.736835, 11.700665, 11.773004, 11.834491, 11.8308735, 11.812789, 11.812789, 11.848958, 11.877893, 11.979167, 12.076823, 12.152778, 12.225116, 12.340857, 12.3878765, 12.525318, 12.641059, 12.7568, 12.894242, 12.984664, 13.0027485, 13.161892, 13.2161455, 13.3933735, 13.454861, 13.556134, 13.70081, 13.722511, 13.859954, 13.946759, 14.084202, 14.203559, 14.344618, 14.42419, 14.568866, 14.58695, 14.702691, 14.825665, 14.963108, 15.024595, 15.1222515, 15.20544, 15.328414, 15.455006, 15.534577, 15.664786, 15.769676, 15.842014, 15.983073, 16.073496, 16.210938, 16.257957, 16.37008, 16.540075, 16.597946, 16.66305, 16.847511, 16.901766, 17.035591, 17.15133, 16.88368, 15.99754, 15.133101, 14.283131, 13.415075, 12.999132, 13.053386, 13.089555, 13.118489, 13.183594, 13.125724, 13.187211, 13.165509, 13.241464, 13.208912, 13.299335, 13.313802, 13.270399, 13.299335, 13.400608, 13.364439, 13.375289, 13.43316, 13.447627, 13.451244, 13.487413, 13.494647, 13.566985, 13.516349, 13.53805, 13.610388, 13.588686, 13.661024, 13.570601, 13.751447, 13.722511, 13.7839985, 13.744213, 13.773149, 13.773149, 13.831018, 13.794849, 13.823785, 13.917824, 13.91059, 13.841869, 14.001013, 13.928675, 13.961226, 13.986546, 14.066117, 14.01548, 14.026331, 14.12037, 14.055266, 14.149305, 14.10952, 14.1746235, 14.185474, 14.26143, 14.286748, 14.27228, 14.283131, 14.337384, 14.337384, 14.398871, 14.373553, 14.416956, 14.391638, 14.496528, 14.492911, 14.492911, 14.536314, 14.550781, 14.5652485, 14.579717, 14.623119, 14.64482, 14.623119, 14.637587, 14.684607, 14.717158, 14.782263, 14.746094, 14.728009, 14.829283, 14.89077, 14.898004, 14.916088, 14.934173, 14.934173, 14.992043, 14.999276, 15.006511, 15.049913, 15.107783, 15.118634, 15.158421, 15.143952, 15.162037, 15.198206, 15.165654, 15.219908, 15.295862, 15.259693, 15.248842, 15.350116, 15.382668, 15.389901, 15.4296875, 15.400752, 15.462239, 15.47309, 15.487557, 15.563513, 17.353878, 19.889322, 22.30541, 24.833622, 27.34375, 29.78154, 32.320602, 34.776474, 37.30107, 39.803963, 42.332176, 42.306858, 38.964844, 36.433014, 33.995224, 31.488716, 29.003906, 26.450377, 24.005354, 21.538628, 18.995949, 16.53284, 14.029948, 13.237847, 13.201678, 13.183594, 13.154658, 13.154658, 13.147425, 13.132957, 13.078704, 13.042535, 13.035301, 13.006366, 13.035301, 12.973814, 12.966579, 12.854456, 12.86169, 12.850839, 12.821904, 12.792969, 12.796586, 12.771267, 12.771267, 12.771267, 12.65191, 12.630208, 12.673611, 12.662761, 12.608507, 12.637443, 12.550636, 12.554254, 12.568721, 12.474682, 12.528935, 12.39511, 12.39511, 12.3878765, 12.402344, 12.3878765, 12.311921, 12.264901, 12.282986, 12.286603, 12.246818, 12.275752, 12.217882, 12.160011, 12.170862, 12.160011, 12.145544, 12.094908, 12.062355, 12.004485, 12.029803, 11.990017, 12.000868, 11.946614, 11.932147, 11.888744, 11.859809, 11.899595, 11.874276, 11.812789, 11.841724, 11.841724, 11.769386, 11.780237, 11.762153, 11.675347, 11.642796, 11.668114, 11.67173, 11.610243, 11.581307, 11.584925, 11.537905, 11.534288, 11.555989, 11.498119, 11.411314, 11.422164, 11.436632, 11.389612, 11.34621, 11.349827, 11.378761, 11.281105, 11.302807, 11.226851, 11.252171, 11.226851, 11.201533, 11.121962, 11.165364, 11.150897, 11.114728, 11.067708, 11.056858, 11.071325, 11.024305, 11.017072, 10.970052, 10.955585, 10.959202, 10.948351, 10.883246, 10.912182, 10.865162, 10.901331, 10.796441, 10.760272, 10.763889, 10.73857, 10.720486, 10.828993, 10.73857, 10.622829, 10.677083, 10.6119795, 10.630064, 10.590278, 10.568577, 10.51794, 10.557726, 10.51794, 10.503472, 10.463686, 10.4347515, 10.449219, 10.420283, 10.380498, 10.445601, 10.304543, 10.373264, 10.286458, 10.2683735, 10.304543, 10.246673, 10.188802, 10.264757, 10.174335, 10.152633, 10.159867, 10.120081, 10.138165, 10.09838, 10.120081, 10.083912, 10.000724, 10.047743, 9.993489, 10.018807, 9.971788, 9.950087, 9.881366, 9.89945, 9.892217, 9.856048, 9.863281, 9.856048, 9.837963, 9.758391, 9.765625, 9.78371, 9.751158, 9.704138, 9.696904, 9.635417, 9.660735, 9.642651, 9.617332, 9.610099, 9.548611, 9.552228, 9.523293, 9.497974, 9.458189, 9.490741, 9.505208, 9.472656, 9.443721, 9.411169, 9.458189, 9.403935, 9.364149, 9.335214, 9.324364, 9.320746, 9.3098955, 9.237557, 9.244792, 9.201389, 9.186921, 9.212239, 9.201389, 9.132668, 9.074798, 9.060329, 9.085649, 9.035011, 9.045862, 9.060329, 8.980758, 9.00246, 8.915654, 8.904803, 8.930121, 8.861401, 8.854167, 8.839699, 8.785445, 8.828849, 8.832465, 8.774595, 8.807147, 8.691406, 8.716724, 8.687789, 8.756511, 8.666088, 8.633536, 8.622685, 8.582899, 8.553964, 8.553964, 8.557581, 8.521412, 8.525029, 8.517796, 8.496094, 8.463542, 8.420139, 8.423756, 8.39482, 8.478009, 8.391204, 8.402055, 8.340568, 8.275463, 8.293548, 8.3152485, 8.224827, 8.297164, 8.279079, 8.087384, 7.4363427, 6.7382812, 6.14511, 5.439815, 5.1576967, 5.10706, 5.0708914, 5.114294, 5.0600405, 5.1359954, 5.078125, 5.078125, 5.1215277, 5.0962095, 5.0311055, 5.0998263, 5.0455728, 5.016638, 5.0347223, 5.0311055, 5.04919, 5.013021, 5.038339, 5.038339, 5.00217, 5.027488, 4.976852, 5.00217, 5.013021, 4.9949365, 4.969618, 4.976852, 5.005787, 4.973235, 5.016638, 5.038339, 4.9949365, 4.973235, 5.013021, 4.9913197, 4.9081306, 4.9225984, 4.9334493, 4.900897, 4.864728, 4.864728, 4.9225984, 4.890046, 4.9081306, 4.8791957, 4.9153647, 4.9479165, 4.904514, 4.868345, 4.8864293, 4.8864293, 1.7216436, 2.311198, 3.0381944, 3.656684, 3.9243345, 3.8881655, 3.8809316, 3.942419, 3.9243345, 3.982205, 3.938802, 4.0256076, 3.9858217, 4.0364585, 4.0039062, 4.0364585, 4.0039062, 4.0364585, 4.0690103, 4.1377316, 4.079861, 4.0690103, 4.1341147, 4.1413484, 4.123264, 4.170284, 4.1377316, 4.1666665, 4.1304975, 4.195602, 4.181134, 4.184751, 4.260706, 4.231771, 4.2498555, 4.3113427, 4.3113427, 4.336661, 4.3185763, 4.369213, 4.3547454, 4.3402777, 4.3764467, 4.405382, 4.3909144, 4.405382, 4.448785, 4.408999, 4.4270835, 4.398148, 4.5319734, 4.5319734, 4.5572915, 4.47772, 4.5211225, 4.546441, 4.5247397, 4.5175056, 4.6006947, 4.578993, 4.571759, 4.6043115, 4.622396, 4.662182, 4.662182, 4.7200522, 4.6694155, 4.7055845, 4.763455, 4.723669, 4.7851562, 4.7417536, 4.7453704, 4.748987, 4.788773, 4.796007, 4.788773, 4.8791957, 4.835793, 4.89728, 4.8466434, 4.926215, 4.9225984, 4.8791957, 4.9153647, 4.9189816, 4.9949365, 4.9804688, 5.0094037, 4.9985533, 5.04919, 5.1576967, 5.295139, 5.403646, 5.4470487, 5.530237, 5.6278934, 5.7689524, 5.8774595, 5.9461803, 6.000434, 6.1197915, 6.1957464, 6.311487, 6.4055266, 6.4778647, 6.5827546, 6.651476, 6.752749, 6.893808, 6.9372106, 7.0457177, 7.1506076, 7.1940103, 7.316985, 7.4363427, 7.5665507, 7.5846353, 7.700376, 7.8305845, 7.8993053, 7.96441, 8.076533, 8.105469, 8.300781, 8.369502, 8.4816265, 8.532263, 8.680555, 8.7890625, 8.886719, 8.95544, 9.0494795, 9.168837, 9.248408, 9.313513, 9.469039, 9.465423, 9.6535015, 9.725839, 9.331597, 8.5286455, 7.7256947, 6.929977, 6.0800056, 5.7689524, 5.797888, 5.758102, 5.855758, 5.848524, 5.8412905, 5.83044, 5.8449073, 5.895544, 5.9534144, 5.8810763, 5.9497976, 5.9534144, 5.910012, 5.9932003, 5.9787326, 6.032986, 5.9823494, 6.0583043, 6.047454, 6.061921, 6.047454, 6.1270256, 6.0872397, 6.1306424, 6.174045, 6.1197915, 6.1306424, 6.2319155, 6.188513, 6.2029805, 6.2174478, 6.213831, 6.2355323, 6.25, 6.3440394, 6.2970195, 6.2644677, 6.358507, 6.289786, 6.3331885, 6.3187213, 6.438079, 6.3729744, 6.3729744, 6.427228, 6.4091434, 6.4453125, 6.4561634, 6.492332, 6.4850984, 6.575521, 6.514034, 6.5610533, 6.5574365, 6.5574365, 6.6840277, 6.6225405, 6.640625, 6.61169, 6.741898, 6.6948786, 6.676794, 6.7238135, 6.6731772, 6.792535, 6.7274303, 6.7853007, 6.7599826, 6.778067, 6.778067, 6.7744503, 6.8467884, 6.890191, 6.9372106, 6.850405, 6.922743, 6.9516783, 6.9335938, 6.9480615, 6.9625287, 6.980613, 6.9842305, 7.0095487, 7.027633, 7.103588, 7.0638022, 7.0746527, 7.1144385, 7.13614, 7.143374, 7.8197336, 10.300926, 12.771267, 15.295862, 17.798756, 20.283566, 22.793692, 25.296585, 27.734375, 30.197483, 32.736546, 35.232204, 37.702545, 40.227142, 40.165653, 37.08044, 34.599247, 32.08912, 29.564526, 27.155672, 24.631077, 22.128183, 19.56742, 17.126013, 14.626736, 12.163629, 9.642651, 7.1289062, 5.4108796, 5.4144964, 5.36386, 5.353009, 5.3891783, 5.3023725, 5.287905, 5.287905, 5.3240743, 5.2336516, 5.2372684, 5.280671, 5.219184, 5.219184, 5.1359954, 5.219184, 5.179398, 5.143229, 5.143229, 5.1685476, 5.074508, 5.0925927, 5.0455728, 5.0962095, 5.027488, 4.9551506, 5.0347223, 5.0094037, 5.027488, 4.9949365, 4.9804688, 4.926215, 4.9117475, 4.962384, 4.89728, 4.875579, 4.890046, 4.8466434, 4.7743053, 4.79239, 4.8213253, 4.8177085, 4.83941, 4.796007, 4.727286, 4.716435, 4.6802664, 4.7019677, 4.6875, 4.6694155, 4.647714, 4.626013, 4.651331, 4.586227, 4.636863, 4.626013, 4.539207, 4.499421, 4.560909, 4.5428243, 4.53559, 4.5319734, 4.4560184, 4.474103, 4.474103, 4.448785, 4.5211225, 4.4632525, 4.4162326, 4.3836803, 4.336661, 4.3511286, 4.296875, 4.3185763, 4.3511286, 4.3149595, 4.3041086, 4.347512, 4.2643228, 4.271557, 4.260706, 4.235388, 4.3041086, 4.1739006, 4.188368, 4.195602, 4.159433, 4.1521993, 4.119647, 4.119647, 4.108796, 4.1015625, 4.05816, 4.123264, 4.0726275, 4.083478, 3.9605036, 4.0039062, 4.007523, 4.0256076, 3.9858217, 3.8990161, 3.9568865, 3.9171007, 3.9641204, 3.9207175, 3.9026332, 3.8773148, 3.8447628, 3.8483796, 3.8447628, 3.8266783, 3.830295, 3.804977, 3.7760417, 3.7507234, 3.7000868, 3.7543402, 3.7181714, 3.7000868, 3.69647, 3.685619, 3.6892362, 3.725405, 3.6639178, 3.6385996, 3.5879629, 3.6385996, 3.5807292, 3.59158, 3.5264757, 3.5083911, 3.5228589, 3.5300925, 3.4975405, 3.5011575, 3.4324362, 3.4252026, 3.5011575, 3.4324362, 3.410735, 3.4360533, 3.3962674, 3.374566, 3.370949, 3.3673322, 3.3528645, 3.3166957, 3.378183, 3.302228, 3.2841434, 3.294994, 3.233507, 3.2732928, 3.2045717, 3.226273, 3.1864872, 3.2045717, 3.2118056, 3.1394675, 3.157552, 3.161169, 3.1358507, 3.1286168, 3.1286168, 3.0454283, 3.0635128, 3.0996816, 3.0454283, 3.049045, 3.049045, 3.023727, 3.0092592, 2.9513888, 2.9513888, 2.983941, 2.980324, 2.9296875, 2.911603, 2.8573496, 2.8645833, 2.9188368, 2.911603, 2.8175638, 2.8537326, 2.842882, 2.8320312, 2.7958622, 2.7777777, 2.8139467, 2.734375, 2.7199075, 2.7596934, 2.7162905, 2.698206, 2.7416089, 2.6945891, 2.6801214, 2.6728878, 2.6367188, 2.629485, 2.6801214, 2.6367188, 2.6150174, 2.5752316, 2.564381, 2.55353, 2.5788484, 2.5426793, 2.4920428, 2.5282118, 2.5065105, 2.5028934, 2.4775753, 2.44864, 2.4088542, 2.4233217, 2.5065105, 2.3980036, 2.445023, 2.3582175, 2.4233217, 2.3618345, 2.376302, 2.3654513, 2.2858796, 2.3184316, 2.23886, 2.3365161, 2.275029, 2.2605612, 2.1918402, 2.2280092, 1.634838, 0.9765625, 0.30020255, 3.4432871, 5.0455728, 5.0998263, 5.10706, 5.0853586, 5.1613135, 5.117911, 5.128762, 5.0925927, 5.143229, 5.0600405, 5.0708914, 5.1649303, 5.128762, 5.114294, 5.103443, 5.1576967, 5.183015, 5.117911, 5.1576967, 5.179398, 5.1649303, 5.0708914, 5.1251445, 5.215567, 5.179398, 5.2119503, 5.1721644, 5.204716, 5.150463, 5.204716, 5.179398, 5.190249, 5.1974826, 5.2445025, 5.2408853, 5.1757812, 5.251736, 5.280671, 5.2445025, 5.255353, 5.2842884, 5.2408853, 5.280671, 5.2445025, 5.2336516, 5.2987556, 5.230035, 5.2698207, 5.31684, 5.3783274, 5.3385415, 5.2987556, 5.287905, 5.3132234, 5.2770543, 5.3747106, 5.3132234, 5.4000287, 5.353009, 5.3096066, 5.6315103, 6.3368053, 6.969763, 7.60272, 8.282697, 8.427373, 8.405671, 8.445457, 8.456307, 8.423756, 8.510561, 8.539496, 8.564815, 8.496094, 8.59375, 8.600984, 8.619068, 8.557581, 8.691406, 8.669704, 8.691406, 8.738426, 8.637153, 8.763744, 8.781829, 8.796296, 8.785445, 8.80353, 8.843316, 8.854167, 8.875868, 8.843316, 8.908421, 8.937355, 8.9192705, 9.006077, 8.959057, 8.998842, 8.973524, 9.016927, 9.031395, 9.031395, 8.998842, 9.085649, 9.063947, 9.154369, 9.186921, 9.161603, 9.273726, 9.201389, 9.226707, 9.233941, 9.248408, 9.248408, 9.338831, 9.338831, 9.349682, 9.302662, 9.364149, 9.447338, 9.367766, 9.454572, 9.385851, 9.42202, 9.476274, 9.490741, 9.505208, 9.505208, 9.602864, 9.555845, 9.544994, 9.588397, 9.628182, 9.664351, 9.628182, 9.660735, 9.682436, 9.729456, 9.707755, 9.73669, 9.740307, 9.823495, 9.805411, 9.798177, 9.823495, 9.866899, 9.881366, 9.85243, 9.975405, 10.007957, 9.95732, 10.029658, 10.185185, 10.206886, 10.315393, 10.467303, 10.554109, 10.691551, 10.756655, 10.789207, 10.966435, 11.067708, 11.161748, 11.205151, 11.338976, 11.472801, 11.555989, 11.603009, 11.715133, 11.794704, 11.924913, 12.040654, 12.131077, 12.203414, 12.355324, 12.384259, 12.507234, 12.60489, 12.648293, 12.800202, 12.9557295, 13.042535, 13.078704, 13.165509, 13.32827, 13.404224, 13.527199, 13.58507, 13.726129, 13.820168, 13.968461, 13.990162, 14.134838, 14.21441, 14.279514, 14.362702, 14.532697, 14.619502, 14.7316265, 14.840133, 14.923322, 14.623119, 13.798467, 12.9557295, 12.160011, 11.382379, 11.020689, 11.053241, 11.121962, 11.107494, 11.143663, 11.121962, 11.150897, 11.14728, 11.219618, 11.190682, 11.183449, 11.223235, 11.302807, 11.295573, 11.255787, 11.364294, 11.317274, 11.375145, 11.3932295, 11.418548, 11.4402485, 11.469184, 11.436632, 11.494502, 11.494502, 11.588542, 11.555989, 11.559607, 11.603009, 11.617476, 11.617476, 11.704283, 11.693432, 11.678964, 11.715133, 11.744068, 11.773004, 11.758536, 11.816406, 11.809173, 11.848958, 11.910445, 11.950232, 11.874276, 11.932147, 11.924913, 11.968316, 11.979167, 12.004485, 12.037037, 12.000868, 12.123842, 12.105758, 12.181713, 12.141927, 12.203414, 12.13831, 12.203414, 12.239583, 12.250434, 12.2432, 12.29022, 12.326389, 12.366175, 12.362557, 12.358941, 12.3878765, 12.3878765, 12.424046, 12.405961, 12.485533, 12.528935, 12.528935, 12.528935, 12.54702, 12.554254, 12.615741, 12.619358, 12.626592, 12.662761, 12.6953125, 12.764033, 12.811053, 12.724248, 12.760417, 12.80382, 12.843605, 12.836371, 12.850839, 12.90871, 12.941261, 13.292101, 15.704572, 18.17853, 20.706741, 23.1807, 25.672743, 28.121384, 30.671297, 33.15249, 35.633682, 38.151043, 40.588833, 40.559895, 37.492767, 34.964554, 32.508682, 30.016638, 27.50651, 25.043404, 22.518808, 20.070168, 17.520254, 15.089699, 12.579572, 11.237702, 11.161748, 11.2160015, 11.114728, 11.100261, 11.121962, 11.096643, 11.085793, 11.031539, 11.024305, 11.056858, 10.951967, 11.020689, 10.944734, 10.912182, 10.901331, 10.87963, 10.8253765, 10.803675, 10.789207, 10.73857, 10.745805, 10.781974, 10.706018, 10.724103, 10.593895, 10.673467, 10.6807, 10.572193, 10.554109, 10.579427, 10.503472, 10.521557, 10.52879, 10.463686, 10.445601, 10.46007, 10.532408, 10.420283, 10.35518, 10.322627, 10.326244, 10.3515625, 10.286458, 10.250289, 10.243055, 10.228588, 10.2213545, 10.181568, 10.206886, 10.192419, 10.083912, 10.112847, 10.083912, 10.054976, 10.047743, 10.007957, 10.007957, 9.964555, 9.982639, 9.986256, 9.924768, 9.89945, 9.892217, 9.848814, 9.837963, 9.884983, 9.801794, 9.780092, 9.780092, 9.754774, 9.725839, 9.725839, 9.711371, 9.693287, 9.6535015, 9.617332, 9.628182, 9.599248, 9.566695, 9.610099, 9.57393, 9.508825, 9.4871235, 9.443721, 9.414786, 9.43287, 9.382234, 9.382234, 9.360533, 9.324364, 9.338831, 9.306279, 9.378617, 9.244792, 9.215857, 9.2628765, 9.291811, 9.186921, 9.183305, 9.190538, 9.194155, 9.147136, 9.067564, 9.035011, 9.009693, 9.103733, 8.991609, 9.009693, 9.009693, 8.991609, 9.027778, 8.933739, 8.8722515, 8.933739, 8.865017, 8.875868, 8.843316, 8.7890625, 8.843316, 8.74566, 8.713108, 8.767361, 8.7058735, 8.687789, 8.673322, 8.7058735, 8.600984, 8.597367, 8.604601, 8.600984, 8.575665, 8.532263, 8.532263, 8.521412, 8.553964, 8.5286455, 8.478009, 8.4816265, 8.470776, 8.409288, 8.351418, 8.308015, 8.362268, 8.3152485, 8.3152485, 8.297164, 8.293548, 8.213976, 8.206742, 8.199508, 8.224827, 8.192274, 8.17419, 8.18504, 8.134404, 8.101851, 8.065682, 8.080151, 8.065682, 8.065682, 8.025897, 7.9716434, 8.036748, 7.9318576, 7.939091, 7.949942, 7.913773, 7.9029226, 7.8703704, 7.884838, 7.8956885, 7.837818, 7.8052664, 7.747396, 7.7582464, 7.7256947, 7.7546296, 7.703993, 7.6931424, 7.7293115, 7.6678243, 7.6171875, 7.5882525, 7.6497397, 7.5810184, 7.573785, 7.5810184, 7.530382, 7.5520835, 7.5050635, 7.486979, 7.472512, 7.5014467, 7.396557, 7.382089, 7.458044, 7.360388, 7.3423033, 7.349537, 7.309751, 7.3025174, 7.248264, 7.306134, 7.269965, 7.2265625, 7.1903934, 7.157841, 7.2012444, 7.139757, 7.168692, 7.1108217, 7.081887, 7.0746527, 7.0999713, 7.0457177, 7.1759257, 7.027633, 7.03125, 6.9878473, 6.9733796, 7.0131655, 6.929977, 6.8757234, 6.8974247, 6.857639, 6.8467884, 6.8865743, 6.8106194, 6.7599826, 6.792535, 6.814236, 6.792535, 6.2970195, 5.6351275, 4.875579, 4.257089, 3.6639178, 3.7073207, 3.69647, 3.6385996, 3.692853, 3.685619, 3.660301, 3.6639178, 3.6385996, 3.656684, 3.7181714, 3.685619, 3.6422164, 3.6277487, 3.620515, 3.6458333, 3.6385996, 3.5951967, 3.584346, 3.6313658, 3.5988138, 3.5879629, 3.5807292, 3.5879629, 3.5554109, 3.5879629, 3.59158, 3.551794, 3.5300925, 3.6060474, 3.5554109, 3.5300925, 3.5409434, 3.5264757, 3.5047743, 3.5192418, 3.5083911, 3.5373263, 3.5626447, 3.5011575, 3.5409434, 3.4866898, 3.5662615, 3.5120082, 3.5047743, 3.5192418, 3.4903066, 3.5228589, 3.4866898, 3.4505208, 3.4722223, 3.4649885, 3.446904, 3.4577546, 3.3528645, 3.4939237, 3.4866898, 3.4179688, 3.4215856, 3.4252026, 3.378183, 1.8916377, 4.615162, 4.626013, 4.5645256, 4.6187787, 4.6187787, 4.560909, 4.662182, 4.6296296, 4.6187787, 4.615162, 4.5645256, 4.622396, 4.6079283, 4.658565, 4.683883, 4.622396, 4.6043115, 4.691117, 4.6875, 4.676649, 4.647714, 4.6440973, 4.651331, 4.691117, 4.5898438, 4.6043115, 4.6730323, 4.723669, 4.6332464, 4.6730323, 4.7019677, 4.727286, 4.698351, 4.7019677, 4.6875, 4.6802664, 4.6730323, 4.6802664, 4.716435, 4.6947336, 4.6549478, 4.727286, 4.7345195, 4.738137, 4.727286, 4.788773, 4.7815394, 4.788773, 4.7670717, 4.7706885, 4.799624, 4.738137, 4.738137, 4.8177085, 4.763455, 4.8574944, 4.7815394, 4.7670717, 4.796007, 4.803241, 4.9479165, 5.5917244, 6.2934027, 6.919126, 7.526765, 7.8956885, 7.8920717, 7.8920717, 7.939091, 7.9029226, 7.960793, 7.960793, 7.960793, 7.9788775, 7.96441, 7.9463253, 8.036748, 8.018663, 8.087384, 8.065682, 8.105469, 8.141638, 8.188658, 8.145255, 8.181423, 8.192274, 8.17419, 8.275463, 8.206742, 8.199508, 8.308015, 8.257379, 8.311632, 8.326099, 8.33695, 8.322483, 8.33695, 8.3152485, 8.412905, 8.380353, 8.344184, 8.463542, 8.412905, 8.467158, 8.459925, 8.525029, 8.496094, 8.499711, 8.568432, 8.499711, 8.575665, 8.564815, 8.619068, 8.626302, 8.684173, 8.629919, 8.684173, 8.69864, 8.662471, 8.713108, 8.716724, 8.785445, 8.774595, 8.785445, 8.7890625, 8.79268, 8.846932, 8.825232, 8.904803, 8.890336, 8.930121, 8.987992, 8.973524, 8.944589, 8.933739, 9.07118, 9.01331, 9.038629, 9.020544, 9.056713, 9.07118, 9.038629, 9.125434, 9.1182, 9.103733, 9.190538, 9.139901, 9.215857, 9.244792, 9.226707, 9.284577, 9.302662, 9.400318, 9.519676, 9.602864, 9.696904, 9.801794, 9.870515, 9.94647, 10.058594, 10.174335, 10.275608, 10.380498, 10.456452, 10.568577, 10.698785, 10.745805, 10.836226, 10.944734, 11.078559, 11.085793, 11.248553, 11.367911, 11.458333, 11.530671, 11.621094, 11.700665, 11.841724, 11.92853, 12.029803, 12.152778, 12.207031, 12.344474, 12.377026, 12.518085, 12.637443, 12.713397, 12.811053, 12.883391, 13.064236, 13.089555, 13.22338, 13.292101, 13.436776, 13.527199, 13.610388, 13.718895, 13.820168, 13.932292, 14.001013, 14.073351, 13.943142, 13.136574, 12.380642, 11.563224, 10.662616, 10.199653, 10.206886, 10.275608, 10.264757, 10.257524, 10.271991, 10.282842, 10.322627, 10.402199, 10.3515625, 10.36603, 10.423901, 10.470921, 10.489005, 10.478154, 10.536024, 10.525173, 10.521557, 10.539641, 10.568577, 10.622829, 10.604745, 10.640914, 10.63368, 10.615596, 10.6589985, 10.698785, 10.767506, 10.687934, 10.724103, 10.78559, 10.807292, 10.854311, 10.756655, 10.821759, 10.774739, 10.876013, 10.857928, 10.894097, 10.857928, 10.926649, 10.930266, 10.988136, 11.035156, 11.046007, 11.038774, 11.017072, 11.096643, 11.118345, 11.085793, 11.143663, 11.201533, 11.1943, 11.201533, 11.176215, 11.230469, 11.205151, 11.342592, 11.291956, 11.31004, 11.313658, 11.313658, 11.331742, 11.41493, 11.443866, 11.407697, 11.46195, 11.447483, 11.490886, 11.51982, 11.541522, 11.545139, 11.501736, 11.628327, 11.621094, 11.628327, 11.639178, 11.624711, 11.646412, 11.682581, 11.729601, 11.71875, 11.791088, 11.794704, 11.856193, 11.834491, 11.780237, 11.845342, 11.852575, 11.859809, 11.932147, 12.084057, 14.369936, 16.880064, 19.382957, 21.849682, 24.374277, 26.837385, 29.394531, 31.807003, 34.324364, 36.816406, 39.304832, 41.82581, 41.822193, 38.697193, 36.23047, 33.716724, 31.210215, 28.68562, 26.182726, 23.672598, 21.216724, 18.75, 16.26519, 13.75868, 11.2160015, 10.21412, 10.170717, 10.199653, 10.116464, 10.058594, 10.112847, 10.073061, 10.10923, 10.080296, 9.993489, 10.015191, 10.040509, 9.968171, 9.928386, 9.924768, 9.982639, 9.942853, 9.859664, 9.870515, 9.845197, 9.845197, 9.834346, 9.85243, 9.686053, 9.765625, 9.725839, 9.73669, 9.718605, 9.7005205, 9.671586, 9.628182, 9.613715, 9.599248, 9.508825, 9.519676, 9.508825, 9.47989, 9.530526, 9.505208, 9.4401045, 9.461805, 9.458189, 9.396702, 9.360533, 9.389467, 9.295428, 9.331597, 9.306279, 9.284577, 9.313513, 9.233941, 9.295428, 9.230324, 9.226707, 9.215857, 9.136285, 9.129051, 9.0964985, 9.1182, 9.0964985, 9.056713, 9.085649, 9.042245, 9.016927, 8.998842, 9.006077, 8.959057, 8.995226, 8.933739, 8.886719, 8.868634, 8.868634, 8.886719, 8.861401, 8.825232, 8.846932, 8.723958, 8.7890625, 8.74566, 8.716724, 8.676939, 8.64077, 8.695024, 8.65162, 8.637153, 8.648004, 8.64077, 8.615452, 8.586516, 8.568432, 8.539496, 8.539496, 8.470776, 8.532263, 8.423756, 8.430989, 8.44184, 8.365886, 8.485243, 8.344184, 8.373119, 8.304399, 8.355035, 8.3152485, 8.300781, 8.246528, 8.297164, 8.257379, 8.235677, 8.206742, 8.199508, 8.177807, 8.159722, 8.152489, 8.065682, 8.148871, 8.083767, 8.065682, 8.051215, 8.047599, 8.029514, 8.01143, 7.9824944, 7.9571757, 7.9427085, 7.921007, 7.924624, 7.888455, 7.8956885, 7.8450522, 7.816117, 7.8305845, 7.873987, 7.7944155, 7.7980323, 7.675058, 7.751013, 7.736545, 7.675058, 7.6569734, 7.7329283, 7.664207, 7.6822915, 7.624421, 7.624421, 7.599103, 7.5810184, 7.5774016, 7.533999, 7.494213, 7.548466, 7.4652777, 7.530382, 7.4905963, 7.3893228, 7.411024, 7.3676214, 7.458044, 7.411024, 7.3350697, 7.3314524, 7.313368, 7.309751, 7.3025174, 7.2663484, 7.284433, 7.2374134, 7.233796, 7.244647, 7.219329, 7.132523, 7.143374, 7.143374, 7.096354, 7.0746527, 7.1289062, 7.0638022, 7.1252894, 7.0529513, 7.0638022, 7.027633, 6.9444447, 7.0638022, 6.9769964, 6.9408274, 6.966146, 6.9625287, 6.893808, 6.9625287, 6.890191, 6.890191, 6.8721066, 6.8359375, 6.8033853, 6.7997684, 6.745515, 6.749132, 6.781684, 6.702112, 6.7853007, 6.7382812, 6.7093463, 6.6731772, 6.629774, 6.6478586, 6.589988, 6.6080728, 6.6623263, 6.604456, 6.5502024, 6.5502024, 6.528501, 6.4742475, 6.503183, 6.463397, 6.4561634, 6.430845, 6.4199944, 6.4344616, 6.488715, 6.3946757, 6.391059, 6.311487, 6.351273, 6.3187213, 6.351273, 6.3078704, 6.275318, 6.2825522, 6.300637, 6.2355323, 6.25, 6.1957464, 5.5157695, 4.9189816, 4.235388, 3.6639178, 3.1394675, 3.125, 3.125, 3.092448, 3.0996816, 3.1141493, 3.1141493, 3.1213832, 3.0743635, 3.1032987, 3.092448, 3.1141493, 3.0996816, 3.1286168, 3.0381944, 3.1177661, 3.1539352, 3.0996816, 3.0635128, 3.0779803, 3.1032987, 3.0743635, 3.0309606, 3.02011, 3.0960648, 3.0635128, 3.092448, 3.0418112, 3.0526621, 3.0454283, 3.0707464, 3.0309606, 3.0345776, 3.0273438, 3.0128763, 3.0671296, 3.0020254, 3.0418112, 3.0526621, 2.9911747, 2.983941, 3.016493, 3.0598958, 3.0598958, 3.0418112, 2.9947917, 2.9911747, 3.0020254, 3.023727, 2.9911747, 2.9947917, 3.0056424, 2.9947917, 2.9767072, 2.947772, 2.9694734, 2.9694734, 2.947772, 2.9730902, 3.023727, 0.003616898, 3.8917825, 7.8667536, 10.387732, 10.405816, 10.4347515, 10.358796, 10.4347515, 10.423901, 10.423901, 10.405816, 10.391349, 10.441985, 10.423901, 10.427517, 10.445601, 10.46007, 10.463686, 10.507089, 10.4347515, 10.427517, 10.496239, 10.456452, 10.478154, 10.463686, 10.496239, 10.496239, 10.4817705, 10.416667, 10.499855, 10.51794, 10.525173, 10.532408, 10.489005, 10.507089, 10.532408, 10.496239, 10.52879, 10.590278, 10.507089, 10.550492, 10.543258, 10.561342, 10.604745, 10.590278, 10.57581, 10.601129, 10.554109, 10.543258, 10.57581, 10.604745, 10.666233, 10.640914, 10.604745, 10.6119795, 10.622829, 10.6119795, 10.63368, 10.637298, 10.669849, 10.6589985, 10.626447, 10.6807, 10.912182, 11.490886, 12.087673, 12.807436, 13.472945, 13.718895, 13.733362, 13.75868, 13.827401, 13.834636, 13.878038, 13.8671875, 13.906974, 13.86357, 13.896123, 13.928675, 13.982928, 13.964844, 14.00463, 13.939526, 14.037182, 14.033565, 14.102286, 14.1276045, 14.080585, 14.1276045, 14.102286, 14.171007, 14.156539, 14.1746235, 14.210793, 14.221643, 14.265046, 14.239728, 14.268663, 14.279514, 14.333767, 14.297599, 14.312066, 14.355469, 14.362702, 14.406105, 14.402489, 14.409722, 14.514612, 14.48206, 14.500145, 14.510995, 14.456742, 14.525463, 14.561632, 14.63397, 14.58695, 14.615886, 14.63397, 14.688224, 14.655671, 14.670139, 14.713542, 14.709925, 14.775029, 14.782263, 14.800347, 14.811198, 14.847367, 14.9088545, 14.854601, 14.869068, 14.90162, 14.934173, 14.923322, 14.959491, 14.945024, 15.002893, 15.028212, 15.05353, 15.0390625, 15.071614, 15.060764, 15.075232, 15.143952, 15.140336, 15.165654, 15.172888, 15.194589, 15.212673, 15.237992, 15.230758, 15.274161, 15.292245, 15.259693, 15.436921, 15.47309, 15.56713, 15.704572, 15.809462, 15.925202, 15.99754, 16.040943, 16.229021, 16.29051, 16.413485, 16.45327, 16.594328, 16.735388, 16.771557, 16.945168, 16.974104, 17.086227, 17.126013, 17.256222, 17.386429, 17.520254, 17.563658, 17.690248, 17.82769, 17.914497, 17.939816, 18.051939, 18.171297, 18.254484, 18.381077, 18.525753, 18.612558, 18.663195, 18.757235, 18.898293, 18.981482, 19.089989, 19.245516, 19.288918, 19.433594, 19.560184, 19.599972, 19.62529, 19.806135, 19.896557, 19.979746, 20.120804, 20.225695, 20.330584, 20.272715, 19.480614, 18.565538, 17.856627, 17.006655, 16.485823, 16.44242, 16.550926, 16.456886, 16.540075, 16.56901, 16.554543, 16.608797, 16.597946, 16.659433, 16.71007, 16.724537, 16.735388, 16.677517, 16.728153, 16.735388, 16.861979, 16.796875, 16.83666, 16.847511, 16.854746, 16.912615, 16.876448, 16.959635, 17.006655, 16.934317, 16.988571, 16.988571, 17.01389, 17.089844, 17.158566, 17.078993, 17.158566, 17.122396, 17.205584, 17.227285, 17.24537, 17.216434, 17.238136, 17.31409, 17.30324, 17.364729, 17.346643, 17.433449, 17.4443, 17.415365, 17.386429, 17.404514, 17.45515, 17.509403, 17.534721, 17.574509, 17.574509, 17.545572, 17.603443, 17.635996, 17.668547, 17.730034, 17.733652, 17.730034, 17.766203, 17.831308, 17.798756, 17.849392, 17.824074, 17.914497, 17.892796, 17.939816, 17.943432, 18.00492, 18.019386, 18.041088, 18.055555, 18.023003, 18.091724, 18.149595, 18.124277, 18.185764, 18.214699, 18.17853, 18.2364, 18.258102, 18.27257, 18.315971, 18.315971, 18.381077, 18.359375, 18.370226, 18.471498, 18.48235, 18.467882, 18.4932, 20.554832, 23.021557, 25.56062, 27.987558, 30.50492, 33.062065, 35.467304, 37.94126, 40.46224, 40.505642, 36.4511, 32.461662, 29.644096, 27.083334, 24.660011, 22.063078, 19.632523, 17.111546, 14.594184, 12.149161, 9.8307295, 9.42202, 9.497974, 9.436487, 9.360533, 9.367766, 9.302662, 9.299046, 9.2628765, 9.324364, 9.230324, 9.2628765, 9.201389, 9.248408, 9.161603, 9.139901, 9.129051, 9.129051, 9.053096, 9.082031, 9.038629, 9.01331, 8.987992, 8.95544, 8.940972, 8.940972, 8.9192705, 8.904803, 8.901186, 8.915654, 8.828849, 8.832465, 8.810764, 8.79268, 8.738426, 8.752893, 8.749276, 8.65162, 8.669704, 8.65162, 8.626302, 8.586516, 8.633536, 8.575665, 8.586516, 8.5286455, 8.470776, 8.434607, 8.430989, 8.478009, 8.409288, 8.365886, 8.33695, 8.409288, 8.333333, 8.344184, 8.347801, 8.318866, 8.322483, 8.308015, 8.192274, 8.250145, 8.206742, 8.192274, 8.163339, 8.058449, 8.105469, 8.112702, 8.047599, 8.029514, 8.080151, 8.015046, 8.0078125, 7.91739, 8.015046, 7.9318576, 7.8956885, 7.8993053, 7.8667536, 7.928241, 7.837818, 7.9065394, 7.7690973, 7.837818, 7.7907987, 7.7437787, 7.7437787, 7.740162, 7.664207, 7.7220774, 7.635272, 7.609954, 7.6063366, 7.6280384, 7.573785, 7.5665507, 7.5159144, 7.5014467, 7.4544272, 7.5050635, 7.4761286, 7.425492, 7.4399595, 7.39294, 7.411024, 7.385706, 7.3350697, 7.3350697, 7.3386865, 7.273582, 7.284433, 7.2663484, 7.2301793, 7.2157116, 7.1976275, 7.157841, 7.1940103, 7.1867766, 7.139757, 7.1144385, 7.096354, 7.081887, 7.0638022, 7.034867, 7.060185, 6.9842305, 6.854022, 6.980613, 6.9408274, 6.929977, 6.904659, 6.9118924, 6.82147, 6.828704, 6.817853, 6.778067, 6.7961516, 6.7310476, 6.7853007, 6.778067, 6.702112, 6.665943, 6.680411, 6.629774, 6.579138, 6.6225405, 6.6550927, 6.5863714, 6.640625, 6.5502024, 6.5610533, 6.514034, 6.467014, 6.4814816, 6.4959493, 6.45978, 6.430845, 6.391059, 6.35489, 6.391059, 6.358507, 6.362124, 6.35489, 6.35489, 6.289786, 6.25, 6.1921296, 6.239149, 6.221065, 6.1921296, 6.1704283, 6.1306424, 6.1631947, 6.1306424, 6.112558, 6.141493, 6.069155, 6.0149016, 6.0257525, 6.0149016, 5.9136286, 5.996817, 5.964265, 5.920862, 5.964265, 5.862992, 5.9136286, 5.870226, 5.8521414, 5.834057, 5.8521414, 5.808738, 5.794271, 5.797888, 5.7725697, 5.7038484, 5.721933, 5.6893806, 5.6532116, 5.721933, 5.67853, 5.6387444, 5.6025753, 5.5664062, 5.5627894, 5.5013022, 5.5483217, 5.4832177, 5.497685, 5.497685, 5.4615164, 5.479601, 5.443432, 5.4361978, 5.392795, 5.3819447, 5.3710938, 5.327691, 5.255353, 5.3132234, 5.2408853, 5.186632, 5.291522, 5.2481194, 5.2372684, 5.2372684, 5.2010994, 5.1974826, 5.1721644, 5.1757812, 5.15408, 5.15408, 5.0962095, 4.9153647, 4.2426214, 3.584346, 2.983941, 2.3039641, 2.0182292, 1.9675926, 1.9929109, 2.0073786, 2.0146122, 1.9748263, 1.9856771, 1.9024885, 1.9712095, 1.8952546, 1.9675926, 1.9748263, 1.9241898, 1.9567419, 1.9458913, 1.9422743, 1.9748263, 1.8735533, 1.9024885, 1.9205729, 1.9241898, 1.9133391, 1.880787, 1.9350405, 1.9567419, 1.8590857, 1.9024885, 1.8880209, 1.8373842, 1.8590857, 1.884404, 1.8699363, 1.8265336, 1.8229166, 1.812066, 1.8554688, 1.8554688, 1.848235, 1.848235, 1.8590857, 1.8265336, 1.775897, 1.8446181, 1.8192998, 1.7903646, 1.8301505, 1.8554688, 1.7903646, 1.739728, 1.8012153, 1.7614294, 1.808449, 1.775897, 1.7469618, 1.7505788, 1.8012153, 1.7650462, 1.7722801, 1.7433449, 1.775897, 2.665654, 6.741898, 6.904659, 6.915509, 6.980613, 6.9625287, 6.8612556, 6.958912, 6.904659, 6.8721066, 6.922743, 6.9372106, 6.929977, 6.955295, 6.9372106, 6.87934, 6.904659, 6.9625287, 6.966146, 6.922743, 6.9625287, 6.92636, 6.958912, 7.0167823, 6.966146, 7.071036, 6.958912, 7.002315, 6.969763, 6.9769964, 6.9842305, 7.0131655, 7.005932, 7.020399, 7.0999713, 7.067419, 7.0384836, 7.0240164, 7.0167823, 7.0384836, 7.060185, 7.0782695, 7.0999713, 7.071036, 7.139757, 7.0891204, 7.0384836, 7.081887, 7.103588, 7.1614585, 7.1216726, 7.1180553, 7.092737, 7.157841, 7.1542244, 7.13614, 7.1614585, 7.107205, 7.18316, 7.146991, 7.2012444, 7.1940103, 7.1903934, 7.107205, 7.2012444, 7.1506076, 7.18316, 7.179543, 7.1903934, 7.1903934, 7.233796, 7.1940103, 7.2012444, 7.2157116, 7.2012444, 7.204861, 7.2518806, 7.269965, 7.2157116, 7.2229457, 7.244647, 7.2916665, 7.24103, 7.2916665, 7.295284, 7.295284, 7.2627316, 7.2518806, 7.3025174, 7.3025174, 7.306134, 7.24103, 7.2916665, 7.313368, 7.418258, 7.3242188, 7.4001737, 7.284433, 7.349537, 7.3386865, 7.3278356, 7.3784723, 7.313368, 7.425492, 7.3748555, 7.3784723, 7.4074073, 7.3640046, 7.418258, 7.4291086, 7.3640046, 7.4001737, 7.421875, 7.3784723, 7.4399595, 7.45081, 7.4037905, 7.4291086, 7.4001737, 7.4652777, 7.4761286, 7.458044, 7.472512, 7.4761286, 7.5014467, 7.4797454, 7.5014467, 7.4363427, 7.4761286, 7.5014467, 7.5159144, 7.5195312, 7.486979, 7.526765, 7.5448494, 7.533999, 7.5448494, 7.570168, 7.5520835, 7.548466, 7.548466, 7.5557003, 7.562934, 7.559317, 7.5810184, 7.60272, 7.526765, 7.5557003, 7.595486, 7.5882525, 7.6533566, 7.6171875, 7.6171875, 7.6425056, 7.6497397, 7.6280384, 7.6497397, 7.6533566, 7.6822915, 7.6533566, 7.703993, 7.696759, 7.70761, 7.6822915, 7.675058, 7.696759, 7.7582464, 7.7220774, 7.6931424, 7.7220774, 7.7329283, 7.7582464, 7.7546296, 7.7220774, 7.7293115, 7.7582464, 7.7293115, 7.761863, 7.7437787, 7.7256947, 7.7582464, 7.7980323, 7.7944155, 7.772714, 7.8595195, 7.837818, 7.8305845, 7.7980323, 7.877604, 7.837818, 7.8812213, 7.9354744, 7.877604, 7.921007, 7.8812213, 7.9029226, 7.949942, 7.8956885, 7.888455, 7.921007, 7.873987, 7.913773, 7.8920717, 7.924624, 7.939091, 7.9354744, 7.939091, 7.9571757, 7.949942, 7.9716434, 7.96441, 7.9824944, 8.02228, 7.993345, 8.047599, 7.989728, 7.986111, 8.058449, 8.015046, 8.087384, 7.9788775, 8.029514, 8.029514, 8.015046, 8.051215, 8.000579, 8.065682, 8.036748, 8.101851, 8.130787, 8.0910015, 8.098235, 8.087384, 8.109086, 8.134404, 8.072917, 8.130787, 8.152489, 8.159722, 8.159722, 8.141638, 8.181423, 8.152489, 8.134404, 8.18504, 8.156105, 8.253761, 8.210359, 8.206742, 8.286314, 8.250145, 8.264612, 8.239294, 8.250145, 8.264612, 8.257379, 8.28993, 8.28993, 8.260995, 8.2682295, 8.326099, 8.3152485, 8.39482, 8.322483, 8.293548, 8.297164, 8.308015, 8.344184, 8.369502, 8.333333, 8.412905, 8.39482, 8.402055, 8.402055, 8.467158, 8.412905, 8.412905, 8.420139, 8.423756, 8.463542, 8.456307, 8.449074, 8.391204, 8.53588, 8.459925, 8.496094, 8.48886, 8.430989, 8.532263, 8.510561, 8.474392, 8.53588, 8.525029, 8.582899, 8.525029, 8.532263, 8.550347, 8.770978, 11.060474, 13.581452, 16.04456, 18.518518, 21.097366, 23.53154, 26.016348, 28.468605, 31.011284, 33.52141, 35.991753, 38.43316, 40.91797, 40.99754, 37.7785, 35.380497, 32.816116, 30.349392, 27.81033, 25.347221, 22.858797, 20.413773, 17.86386, 15.350116, 12.91956, 10.376881, 7.96441, 6.8250866, 6.8612556, 6.8106194, 6.8359375, 6.8395543, 6.8106194, 6.792535, 6.8106194, 6.7744503, 6.7853007, 6.792535, 6.756366, 6.7744503, 6.7274303, 6.7382812, 6.756366, 6.767216, 6.749132, 6.6876445, 6.7635994, 6.7708335, 6.7093463, 6.702112, 6.741898, 6.691262, 6.640625, 6.6948786, 6.6333914, 6.640625, 6.604456, 6.651476, 6.640625, 6.6478586, 6.600839, 6.5936055, 6.6080728, 6.5863714, 6.5863714, 6.6080728, 6.6225405, 6.6189237, 6.579138, 6.615307, 6.6080728, 6.5610533, 6.6225405, 6.528501, 6.5502024, 6.524884, 6.492332, 6.528501, 6.5104165, 6.532118, 6.4453125, 6.488715, 6.4489293, 6.488715, 6.4778647, 6.4706306, 6.463397, 6.40191, 6.4344616, 6.4453125, 6.4416957, 6.4489293, 6.387442, 6.4091434, 6.423611, 6.40191, 6.427228, 6.427228, 6.3946757, 6.376591, 6.45978, 6.3729744, 6.351273, 6.2970195, 6.3838253, 6.358507, 6.325955, 6.3331885, 6.289786, 6.322338, 6.3693576, 6.3295717, 6.2934027, 6.2825522, 6.3042536, 6.325955, 6.184896, 6.260851, 6.2644677, 6.2970195, 6.2174478, 6.2319155, 6.1921296, 6.25, 6.2427664, 6.2029805, 6.210214, 6.199363, 6.239149, 6.184896, 6.213831, 6.1957464, 6.1631947, 6.239149, 6.1559606, 6.1559606, 6.2065973, 6.0872397, 6.1668115, 6.174045, 6.148727, 6.101707, 6.188513, 6.1595774, 6.069155, 6.148727, 6.112558, 6.0944734, 6.0836225, 6.047454, 6.0836225, 6.061921, 6.09809, 6.0872397, 6.061921, 6.1197915, 6.0655384, 6.061921, 6.0185184, 6.0944734, 6.047454, 6.032986, 6.04022, 6.007668, 5.985966, 6.007668, 6.0221353, 5.985966, 5.960648, 5.996817, 5.964265, 5.975116, 6.0293694, 6.0221353, 5.9497976, 5.9570312, 5.964265, 6.0040507, 5.931713, 5.9136286, 5.9497976, 5.924479, 5.9425635, 5.9280963, 5.9136286, 5.8810763, 5.870226, 5.8810763, 5.8412905, 5.9280963, 5.8449073, 5.8449073, 5.8774595, 5.8376737, 5.823206, 5.8810763, 5.855758, 5.855758, 5.797888, 5.8123555, 5.8738427, 5.7761865, 5.7725697, 5.8376737, 5.78342, 5.743634, 5.808738, 5.732784, 5.8051214, 5.7761865, 5.747251, 5.78342, 5.743634, 5.8015046, 5.743634, 5.7364006, 5.747251, 5.7400174, 5.7906537, 5.732784, 5.671296, 5.7400174, 5.6640625, 5.6893806, 5.7038484, 5.656829, 5.7146993, 5.656829, 5.649595, 5.6640625, 5.642361, 5.649595, 5.711082, 5.6676793, 5.6893806, 5.6604457, 5.6315103, 5.642361, 5.6351275, 5.6532116, 5.5989585, 5.6387444, 5.5917244, 5.5989585, 5.5881076, 5.584491, 5.617043, 5.642361, 5.5664062, 5.570023, 5.5230036, 5.62066, 5.580874, 5.5555553, 5.584491, 5.5664062, 5.544705, 5.5374713, 5.5555553, 5.5266204, 5.5374713, 5.580874, 5.5157695, 5.5483217, 5.580874, 5.497685, 5.5013022, 5.497685, 5.5230036, 5.504919, 5.497685, 5.494068, 5.443432, 5.504919, 5.472367, 5.4615164, 5.472367, 5.4506655, 5.457899, 5.3855615, 5.3493924, 5.4144964, 5.4217305, 5.4217305, 5.403646, 5.396412, 5.3855615, 5.428964, 5.3855615, 5.4253473, 5.3819447, 5.3819447, 5.3240743, 5.36386, 5.3493924, 5.360243, 5.3855615, 5.353009, 5.3891783, 5.367477, 5.3747106, 5.3783274, 5.342159, 5.3023725, 5.3385415, 5.2625866, 5.266204, 5.31684, 5.320457, 5.3132234, 5.367477, 5.31684, 5.2372684, 5.295139, 5.2842884, 5.2734375, 5.251736, 5.2698207, 5.2698207, 5.2010994, 5.215567, 5.251736, 5.215567, -0.01808449, 2.0688658, 2.7307582, 3.3600984, 3.8519964, 3.9134839, 3.9026332, 3.8953993, 3.9171007, 3.9568865, 3.9568865, 3.9858217, 4.0039062, 4.018374, 3.9677372, 4.01114, 4.007523, 4.0509257, 4.021991, 4.079861, 4.184751, 4.181134, 4.094329, 4.1304975, 4.1413484, 4.191985, 4.1739006, 4.1775174, 4.170284, 4.2173033, 4.2064524, 4.271557, 4.2100697, 4.195602, 4.2896414, 4.271557, 4.32581, 4.307726, 4.300492, 4.296875, 4.333044, 4.401765, 4.3655963, 4.3511286, 4.3800635, 4.3945312, 4.445168, 4.434317, 4.37283, 4.5030384, 4.448785, 4.4524016, 4.5536747, 4.510272, 4.5645256, 4.546441, 4.575376, 4.575376, 4.5970774, 4.5645256, 4.5898438, 4.6296296, 4.622396, 4.658565, 4.6694155, 4.626013, 4.647714, 4.6694155, 4.7092013, 4.691117, 4.7417536, 4.7200522, 4.7345195, 4.814091, 4.8104744, 4.8828125, 4.799624, 4.8538775, 4.8719616, 4.824942, 4.9081306, 4.8936634, 4.951534, 4.9442997, 4.969618, 4.9840856, 4.9479165, 5.041956, 4.9985533, 5.027488, 5.00217, 5.1215277, 5.25897, 5.356626, 5.418113, 5.494068, 5.5989585, 5.6966147, 5.78342, 5.870226, 5.9895835, 6.047454, 6.188513, 6.275318, 6.3440394, 6.4850984, 6.600839, 6.6550927, 6.749132, 6.781684, 6.8757234, 7.0638022, 7.132523, 7.2265625, 7.2880497, 7.360388, 7.4797454, 7.559317, 7.66059, 7.7690973, 7.863137, 7.9716434, 8.083767, 8.1380205, 8.210359, 8.358651, 8.373119, 8.564815, 8.666088, 8.749276, 8.79268, 8.940972, 9.024161, 9.125434, 9.205006, 9.280961, 9.414786, 9.501592, 9.58478, 9.682436, 9.740307, 8.868634, 8.083767, 7.269965, 6.463397, 5.7689524, 5.8123555, 5.859375, 5.855758, 5.870226, 5.8919272, 5.8919272, 5.895544, 5.975116, 6.011285, 5.9570312, 6.0149016, 6.0040507, 6.072772, 6.076389, 6.069155, 6.0944734, 6.1306424, 6.199363, 6.1704283, 6.1631947, 6.184896, 6.199363, 6.213831, 6.2644677, 6.2717013, 6.3042536, 6.322338, 6.365741, 6.3440394, 6.3838253, 6.3802085, 6.4561634, 6.4091434, 6.4489293, 6.45978, 6.528501, 6.5067997, 6.532118, 6.528501, 6.589988, 6.5936055, 6.5719037, 6.5936055, 6.651476, 6.6731772, 6.702112, 6.712963, 6.7201967, 6.7093463, 6.828704, 6.7961516, 6.7853007, 6.8395543, 6.857639, 6.8974247, 6.8757234, 6.919126, 6.9516783, 6.9335938, 6.929977, 7.0167823, 7.0240164, 6.9733796, 7.056568, 7.042101, 7.168692, 7.146991, 7.1144385, 7.143374, 7.1650753, 7.1506076, 7.212095, 7.2157116, 7.2591147, 7.244647, 7.2916665, 7.309751, 7.2916665, 7.360388, 7.4001737, 7.3386865, 7.39294, 7.4146414, 7.4652777, 7.4544272, 7.483362, 7.494213, 7.4652777, 7.573785, 7.631655, 7.609954, 9.523293, 11.97555, 14.507379, 16.948784, 19.509548, 21.96904, 24.4864, 26.938658, 29.47772, 31.911892, 34.3967, 36.9647, 39.373554, 41.858364, 41.95602, 38.740597, 36.295574, 33.78183, 31.282553, 28.725405, 26.280382, 23.828125, 21.296297, 18.804253, 16.34838, 13.841869, 11.400463, 8.85055, 6.4489293, 5.9172454, 5.870226, 5.8521414, 5.794271, 5.7725697, 5.7761865, 5.7400174, 5.7291665, 5.707465, 5.6966147, 5.671296, 5.6676793, 5.642361, 5.617043, 5.6025753, 5.577257, 5.4868345, 5.5555553, 5.504919, 5.472367, 5.4506655, 5.439815, 5.3891783, 5.443432, 5.3493924, 5.342159, 5.360243, 5.3819447, 5.31684, 5.331308, 5.295139, 5.2842884, 5.2336516, 5.2336516, 5.1757812, 5.190249, 5.2119503, 5.1106772, 5.0962095, 5.067274, 5.10706, 5.0564237, 5.0600405, 4.9877024, 5.0094037, 4.962384, 4.966001, 4.962384, 4.9189816, 4.929832, 4.875579, 4.904514, 4.8430266, 4.8466434, 4.79239, 4.7743053, 4.7779226, 4.763455, 4.712818, 4.712818, 4.698351, 4.6730323, 4.6296296, 4.6694155, 4.636863, 4.5934606, 4.5572915, 4.5898438, 4.550058, 4.510272, 4.513889, 4.448785, 4.434317, 4.448785, 4.4162326, 4.3836803, 4.3438945, 4.412616, 4.3655963, 4.32581, 4.322193, 4.296875, 4.307726, 4.2643228, 4.2498555, 4.260706, 4.2136865, 4.184751, 4.148582, 4.1666665, 4.1739006, 4.0979457, 4.0509257, 4.1304975, 4.11603, 4.0400753, 4.05816, 4.043692, 3.9930556, 4.0002894, 3.9641204, 3.9134839, 3.9460359, 3.9315684, 3.8664641, 3.8809316, 3.8809316, 3.8628473, 3.870081, 3.765191, 3.8194444, 3.7760417, 3.761574, 3.7760417, 3.7145543, 3.7941263, 3.7217882, 3.768808, 3.7181714, 3.7109375, 3.685619, 3.653067, 3.6711516, 3.6747684, 3.6277487, 3.5951967, 3.653067, 3.5807292, 3.5771122, 3.5662615, 3.5879629, 3.5373263, 3.5264757, 3.4939237, 3.479456, 3.5083911, 3.4975405, 3.4541378, 3.4613714, 3.4288194, 3.446904, 3.3564816, 3.4288194, 3.414352, 3.3854167, 3.3926504, 3.3311632, 3.2769098, 3.3962674, 3.3275464, 3.305845, 3.3094618, 3.2443576, 3.2443576, 3.2913773, 3.200955, 3.1973379, 3.2118056, 3.193721, 3.200955, 3.1394675, 3.0960648, 3.1322339, 3.1286168, 3.0852141, 3.056279, 3.0635128, 3.0743635, 3.0635128, 3.0454283, 3.0092592, 3.0056424, 3.0092592, 2.9622395, 2.9658566, 2.980324, 2.9730902, 2.9333043, 2.9333043, 2.879051, 2.879051, 2.879051, 2.904369, 2.8284144, 2.81033, 2.7813947, 2.8211806, 2.8139467, 2.879051, 2.7596934, 2.7633102, 2.7271411, 2.7596934, 2.7090566, 2.6909723, 2.7235243, 2.6439526, 2.7162905, 2.633102, 2.6367188, 2.6439526, 2.6222513, 2.593316, 2.5499132, 2.6114004, 2.5860822, 2.5173612, 2.5752316, 2.4956598, 2.4920428, 2.5499132, 2.4920428, 2.4703414, 2.481192, 2.419705, 2.4414062, 2.44864, 2.3726852, 2.4016204, 2.419705, 2.34375, 2.4016204, 2.3654513, 2.34375, 2.3220487, 2.307581, 2.3148148, 2.3003473, 2.2967303, 2.2822628, 2.2243924, 2.199074, 1.9965278, 1.3599538, 0.77039933, 4.235388, 6.915509, 6.8323207, 6.8865743, 6.9082756, 6.922743, 6.919126, 6.9335938, 6.922743, 6.929977, 6.9082756, 6.9118924, 6.9372106, 6.966146, 6.9372106, 6.966146, 6.969763, 7.002315, 6.969763, 6.9733796, 6.922743, 6.9480615, 6.9516783, 6.9986978, 6.9625287, 6.966146, 7.0384836, 7.0167823, 7.0167823, 7.060185, 6.9769964, 7.027633, 7.020399, 7.042101, 7.034867, 7.107205, 7.0638022, 7.0529513, 6.995081, 7.0638022, 7.060185, 7.03125, 7.0891204, 7.1289062, 7.0891204, 7.0638022, 7.0638022, 7.042101, 7.056568, 7.1289062, 7.060185, 7.132523, 7.1144385, 7.1216726, 7.1216726, 7.1650753, 7.103588, 7.132523, 7.1252894, 7.1614585, 7.13614, 7.3423033, 7.9824944, 8.629919, 9.302662, 9.993489, 10.250289, 10.275608, 10.239439, 10.315393, 10.304543, 10.362413, 10.340712, 10.380498, 10.441985, 10.427517, 10.405816, 10.449219, 10.478154, 10.445601, 10.499855, 10.543258, 10.550492, 10.550492, 10.546875, 10.590278, 10.619213, 10.640914, 10.622829, 10.619213, 10.684318, 10.706018, 10.745805, 10.7421875, 10.821759, 10.771123, 10.767506, 10.774739, 10.821759, 10.8723955, 10.883246, 10.828993, 10.868779, 10.876013, 10.955585, 10.9375, 10.912182, 10.988136, 10.980903, 11.053241, 11.035156, 11.035156, 11.020689, 11.085793, 11.067708, 11.111111, 11.125579, 11.093026, 11.176215, 11.190682, 11.201533, 11.212384, 11.183449, 11.281105, 11.295573, 11.288339, 11.29919, 11.338976, 11.291956, 11.400463, 11.433015, 11.389612, 11.436632, 11.41493, 11.436632, 11.458333, 11.487268, 11.541522, 11.548756, 11.581307, 11.56684, 11.595776, 11.588542, 11.668114, 11.642796, 11.631945, 11.722367, 11.729601, 11.689815, 11.678964, 11.780237, 11.76577, 11.892361, 11.979167, 12.051505, 12.134693, 12.319155, 12.322772, 12.445746, 12.55787, 12.659143, 12.702546, 12.86169, 12.973814, 13.017217, 13.17636, 13.259548, 13.357204, 13.429543, 13.603154, 13.675492, 13.718895, 13.809318, 14.008246, 14.058883, 14.152923, 14.275897, 14.36632, 14.438658, 14.550781, 14.63397, 14.713542, 14.847367, 14.970342, 15.006511, 15.143952, 15.209057, 15.3464985, 15.476707, 15.5598955, 15.700954, 15.650318, 15.878182, 15.968605, 16.059029, 16.109665, 16.257957, 16.304977, 16.489439, 16.536459, 16.713686, 16.749855, 16.681135, 15.849248, 15.04268, 14.228877, 13.440393, 12.879774, 12.865307, 12.995515, 12.962963, 12.905092, 12.926794, 13.013599, 13.017217, 13.096788, 13.035301, 13.104022, 13.100405, 13.1691265, 13.190827, 13.17636, 13.179976, 13.212529, 13.205296, 13.230614, 13.263165, 13.255932, 13.284867, 13.306568, 13.357204, 13.353588, 13.317419, 13.418693, 13.422309, 13.451244, 13.494647, 13.49103, 13.5597515, 13.53805, 13.595921, 13.621239, 13.624855, 13.646557, 13.624855, 13.697193, 13.726129, 13.718895, 13.7369795, 13.762298, 13.798467, 13.751447, 13.838252, 13.812934, 13.86357, 13.903357, 13.870805, 13.986546, 13.972077, 13.935908, 14.019097, 14.044415, 14.0625, 14.1276045, 14.076967, 14.102286, 14.080585, 14.145689, 14.163774, 14.196325, 14.243345, 14.26143, 14.268663, 14.293982, 14.308449, 14.315682, 14.359086, 14.384404, 14.3880205, 14.637587, 17.12963, 19.545717, 22.106482, 24.594908, 27.02908, 29.542824, 32.00955, 34.49074, 37.01172, 39.50376, 41.923466, 41.927082, 38.925056, 36.342594, 33.778214, 31.369358, 28.884548, 26.425058, 23.969185, 21.45544, 18.927229, 16.536459, 14.026331, 12.742332, 12.666377, 12.641059, 12.684462, 12.572338, 12.579572, 12.594039, 12.514467, 12.478298, 12.471065, 12.521702, 12.416811, 12.413195, 12.3878765, 12.416811, 12.351707, 12.319155, 12.333623, 12.333623, 12.275752, 12.286603, 12.297454, 12.188947, 12.185329, 12.188947, 12.1744795, 12.185329, 12.160011, 12.073206, 12.112992, 12.069589, 12.069589, 11.968316, 12.037037, 11.942998, 11.924913, 11.903212, 11.877893, 11.895978, 11.885127, 11.877893, 11.798322, 11.780237, 11.736835, 11.77662, 11.736835, 11.682581, 11.668114, 11.689815, 11.646412, 11.6536455, 11.621094, 11.574074, 11.61386, 11.490886, 11.541522, 11.548756, 11.443866, 11.505353, 11.469184, 11.436632, 11.3932295, 11.371528, 11.3932295, 11.338976, 11.313658, 11.291956, 11.248553, 11.266638, 11.244936, 11.244936, 11.1943, 11.190682, 11.205151, 11.201533, 11.129195, 11.121962, 11.107494, 11.093026, 11.027923, 11.064092, 11.046007, 11.020689, 10.99537, 10.966435, 10.933883, 10.926649, 10.87963, 10.883246, 10.792824, 10.839844, 10.854311, 10.839844, 10.767506, 10.763889, 10.724103, 10.760272, 10.716869, 10.698785, 10.651765, 10.673467, 10.662616, 10.630064, 10.615596, 10.637298, 10.539641, 10.561342, 10.492621, 10.514323, 10.420283, 10.441985, 10.449219, 10.445601, 10.384114, 10.394965, 10.391349, 10.340712, 10.300926, 10.286458, 10.250289, 10.340712, 10.243055, 10.250289, 10.196036, 10.192419, 10.177952, 10.152633, 10.145399, 10.163484, 10.105614, 10.054976, 10.069445, 10.047743, 9.968171, 10.062211, 9.979022, 10.00434, 9.997107, 9.964555, 9.932002, 9.892217, 9.924768, 9.866899, 9.8307295, 9.812645, 9.765625, 9.743923, 9.780092, 9.751158, 9.74754, 9.704138, 9.628182, 9.689671, 9.660735, 9.613715, 9.635417, 9.620949, 9.559462, 9.516059, 9.544994, 9.606482, 9.483507, 9.505208, 9.447338, 9.490741, 9.4401045, 9.436487, 9.382234, 9.403935, 9.382234, 9.371383, 9.331597, 9.31713, 9.27011, 9.306279, 9.248408, 9.259259, 9.27011, 9.172454, 9.143518, 9.139901, 9.1796875, 9.129051, 9.089265, 9.078414, 9.092882, 9.078414, 9.01331, 9.0494795, 8.973524, 8.980758, 9.024161, 8.959057, 9.00246, 8.908421, 8.857783, 8.861401, 8.854167, 8.80353, 8.861401, 8.760127, 8.85055, 8.817998, 8.734809, 8.731193, 8.702257, 8.723958, 8.734809, 8.6588545, 8.619068, 8.615452, 8.608217, 8.579283, 8.503327, 7.8559027, 7.309751, 6.6333914, 5.964265, 5.530237, 5.541088, 5.5121527, 5.4759836, 5.533854, 5.5013022, 5.494068, 5.5013022, 5.5157695, 5.3855615, 5.4470487, 5.439815, 5.544705, 5.4615164, 5.443432, 5.360243, 5.4000287, 5.432581, 5.4000287, 5.367477, 5.4470487, 5.3710938, 5.4253473, 5.3783274, 5.396412, 5.4470487, 5.3240743, 5.3710938, 5.4108796, 5.4361978, 5.342159, 5.353009, 5.367477, 5.4000287, 5.392795, 5.4108796, 5.3059897, 5.331308, 5.3710938, 5.31684, 5.360243, 5.327691, 5.327691, 5.31684, 5.287905, 5.2228007, 5.3493924, 5.331308, 5.2987556, 5.255353, 5.3096066, 5.287905, 5.266204, 5.266204, 5.2119503, 5.2228007, 5.2408853, 5.2842884, 5.230035, 5.1974826, -0.047019675, 1.5661169, 5.5266204, 6.0583043, 6.0908566, 6.0583043, 6.141493, 6.1161747, 6.069155, 6.1631947, 6.076389, 6.101707, 6.141493, 6.1559606, 6.1595774, 6.112558, 6.1523438, 6.141493, 6.076389, 6.2065973, 6.1270256, 6.1053243, 6.101707, 6.1921296, 6.137876, 6.1812787, 6.137876, 6.174045, 6.1921296, 6.2282987, 6.260851, 6.174045, 6.260851, 6.174045, 6.2065973, 6.224682, 6.2427664, 6.246383, 6.2572336, 6.289786, 6.224682, 6.246383, 6.1812787, 6.2825522, 6.213831, 6.239149, 6.224682, 6.260851, 6.2680845, 6.2680845, 6.3042536, 6.253617, 6.2572336, 6.3295717, 6.246383, 6.3187213, 6.3404226, 6.3404226, 6.311487, 6.2717013, 6.325955, 6.286169, 6.278935, 6.87934, 7.494213, 8.11632, 8.828849, 9.371383, 9.414786, 9.461805, 9.505208, 9.483507, 9.461805, 9.566695, 9.476274, 9.566695, 9.592014, 9.58478, 9.642651, 9.58478, 9.689671, 9.711371, 9.671586, 9.67882, 9.646267, 9.696904, 9.74754, 9.790943, 9.787327, 9.812645, 9.85243, 9.841579, 9.863281, 9.866899, 9.89945, 9.884983, 9.950087, 9.953704, 9.997107, 9.979022, 9.993489, 10.047743, 10.0441265, 10.105614, 10.116464, 10.076678, 10.047743, 10.09838, 10.101996, 10.145399, 10.196036, 10.239439, 10.199653, 10.206886, 10.246673, 10.311776, 10.279224, 10.293693, 10.311776, 10.319011, 10.358796, 10.398582, 10.380498, 10.441985, 10.402199, 10.4817705, 10.409432, 10.478154, 10.445601, 10.590278, 10.507089, 10.590278, 10.536024, 10.56496, 10.583044, 10.648149, 10.608362, 10.695168, 10.6807, 10.698785, 10.771123, 10.716869, 10.807292, 10.756655, 10.818142, 10.8253765, 10.8723955, 10.814526, 10.915798, 10.886864, 10.962818, 10.933883, 10.9375, 11.024305, 11.08941, 11.168982, 11.273871, 11.422164, 11.487268, 11.577691, 11.66088, 11.791088, 11.942998, 12.004485, 12.051505, 12.116609, 12.2432, 12.380642, 12.449364, 12.597656, 12.680845, 12.764033, 12.847222, 12.948495, 13.064236, 13.147425, 13.245081, 13.378906, 13.418693, 13.610388, 13.646557, 13.70081, 13.8671875, 13.925057, 14.087818, 14.160156, 14.275897, 14.355469, 14.43504, 14.510995, 14.680989, 14.756945, 14.832899, 14.966724, 15.046296, 15.154803, 15.292245, 15.389901, 15.455006, 15.5598955, 15.628617, 15.794994, 15.867332, 15.954138, 15.353733, 14.612268, 13.7839985, 13.0027485, 12.123842, 12.076823, 12.087673, 12.094908, 12.09129, 12.120226, 12.203414, 12.178096, 12.160011, 12.203414, 12.250434, 12.268518, 12.311921, 12.3046875, 12.3046875, 12.340857, 12.337239, 12.380642, 12.398726, 12.416811, 12.481915, 12.492766, 12.528935, 12.460214, 12.525318, 12.518085, 12.561487, 12.550636, 12.572338, 12.644676, 12.662761, 12.69893, 12.706163, 12.720631, 12.70978, 12.745949, 12.771267, 12.767651, 12.843605, 12.8255205, 12.86169, 12.87254, 12.879774, 12.944879, 12.966579, 12.915943, 12.962963, 12.97743, 13.042535, 13.053386, 13.107639, 13.118489, 13.132957, 13.1691265, 13.12934, 13.198061, 13.194445, 13.248698, 13.263165, 13.274016, 13.292101, 13.321036, 13.342737, 13.3463545, 13.411458, 13.389757, 13.425926, 13.43316, 13.483796, 13.530816, 13.512732, 13.556134, 13.545283, 13.563368, 13.603154, 13.6067705, 13.697193, 13.671875, 13.715278, 13.722511, 13.733362, 13.762298, 13.827401, 13.776765, 13.859954, 13.870805, 13.899739, 13.914207, 13.91059, 13.943142, 13.91059, 14.001013, 14.9088545, 17.379196, 19.874855, 22.363281, 24.927662, 27.434172, 29.868345, 32.37124, 34.84158, 37.351707, 39.850983, 42.30324, 42.317707, 38.404224, 35.919415, 33.412907, 30.917246, 28.464989, 25.951244, 23.441116, 20.916521, 18.478733, 15.9505205, 13.469329, 11.038774, 10.152633, 10.141783, 10.0911455, 10.087529, 10.101996, 10.058594, 10.033276, 10.00434, 9.997107, 9.89945, 9.950087, 9.950087, 9.942853, 9.870515, 9.845197, 9.801794, 9.8307295, 9.798177, 9.790943, 9.790943, 9.725839, 9.664351, 9.7005205, 9.704138, 9.624566, 9.664351, 9.58478, 9.559462, 9.563079, 9.544994, 9.512443, 9.541377, 9.4871235, 9.454572, 9.425636, 9.447338, 9.396702, 9.382234, 9.360533, 9.346065, 9.342448, 9.331597, 9.3098955, 9.288195, 9.212239, 9.241175, 9.172454, 9.215857, 9.168837, 9.154369, 9.132668, 9.092882, 9.027778, 9.092882, 9.024161, 8.984375, 8.987992, 8.948206, 8.908421, 8.937355, 8.875868, 8.893952, 8.861401, 8.854167, 8.828849, 8.832465, 8.817998, 8.756511, 8.785445, 8.770978, 8.709491, 8.655237, 8.74566, 8.6588545, 8.648004, 8.626302, 8.644386, 8.579283, 8.586516, 8.485243, 8.532263, 8.452691, 8.5286455, 8.492476, 8.445457, 8.39482, 8.420139, 8.387587, 8.39482, 8.351418, 8.347801, 8.318866, 8.326099, 8.224827, 8.260995, 8.217592, 8.188658, 8.192274, 8.217592, 8.098235, 8.083767, 8.0910015, 8.065682, 8.065682, 8.051215, 8.051215, 8.076533, 8.015046, 7.9716434, 7.953559, 7.9354744, 7.91739, 7.913773, 7.913773, 7.884838, 7.808883, 7.787182, 7.7907987, 7.8197336, 7.8197336, 7.761863, 7.7582464, 7.700376, 7.7148438, 7.6822915, 7.685909, 7.6461225, 7.6208043, 7.570168, 7.5882525, 7.5882525, 7.5050635, 7.562934, 7.533999, 7.526765, 7.4688945, 7.472512, 7.49783, 7.421875, 7.425492, 7.349537, 7.4037905, 7.3531537, 7.3748555, 7.306134, 7.3314524, 7.3025174, 7.313368, 7.2012444, 7.2229457, 7.295284, 7.248264, 7.172309, 7.172309, 7.1614585, 7.13614, 7.0855036, 7.0746527, 7.0891204, 7.0493345, 7.071036, 7.0167823, 6.966146, 6.9516783, 6.9516783, 6.9118924, 6.922743, 6.8684897, 6.8757234, 6.8250866, 6.8757234, 6.8684897, 6.8033853, 6.7997684, 6.781684, 6.6876445, 6.756366, 6.6948786, 6.6948786, 6.7274303, 6.6731772, 6.680411, 6.6587095, 6.6225405, 6.5863714, 6.604456, 6.575521, 6.5863714, 6.5538197, 6.5212674, 6.4742475, 6.499566, 6.4489293, 6.4344616, 6.4814816, 6.35489, 6.358507, 6.362124, 6.3368053, 6.311487, 6.358507, 6.2717013, 6.289786, 6.2572336, 6.224682, 6.213831, 6.2355323, 6.184896, 6.184896, 6.1812787, 6.09809, 6.1161747, 6.137876, 6.112558, 6.0872397, 6.0257525, 6.0293694, 6.032986, 6.101707, 5.964265, 5.9787326, 5.9497976, 5.964265, 5.910012, 5.910012, 5.862992, 5.9172454, 5.834057, 5.8268228, 5.754485, 5.8376737, 5.787037, 5.7255497, 5.0311055, 4.4958043, 3.8664641, 3.1539352, 2.6511862, 2.6692708, 2.6475694, 2.6692708, 2.7379918, 2.6620371, 2.6837385, 2.6692708, 2.6692708, 2.6114004, 2.6367188, 2.6620371, 2.5788484, 2.6367188, 2.6186342, 2.6150174, 2.6077836, 2.6077836, 2.596933, 2.589699, 2.557147, 2.589699, 2.629485, 2.5788484, 2.6041667, 2.6186342, 2.5499132, 2.5607638, 2.5282118, 2.5354457, 2.589699, 2.6041667, 2.524595, 2.5028934, 2.4739583, 2.4956598, 2.513744, 2.524595, 2.5028934, 2.524595, 2.5065105, 2.5028934, 2.513744, 2.4594908, 2.4594908, 2.419705, 2.4739583, 2.5282118, 2.4414062, 2.4269388, 2.5028934, 2.4377894, 2.4594908, 2.4414062, 2.3943865, 2.4631076, 2.5028934, 2.445023, 2.4305556, 2.4377894, 0.0];
END_VAR
